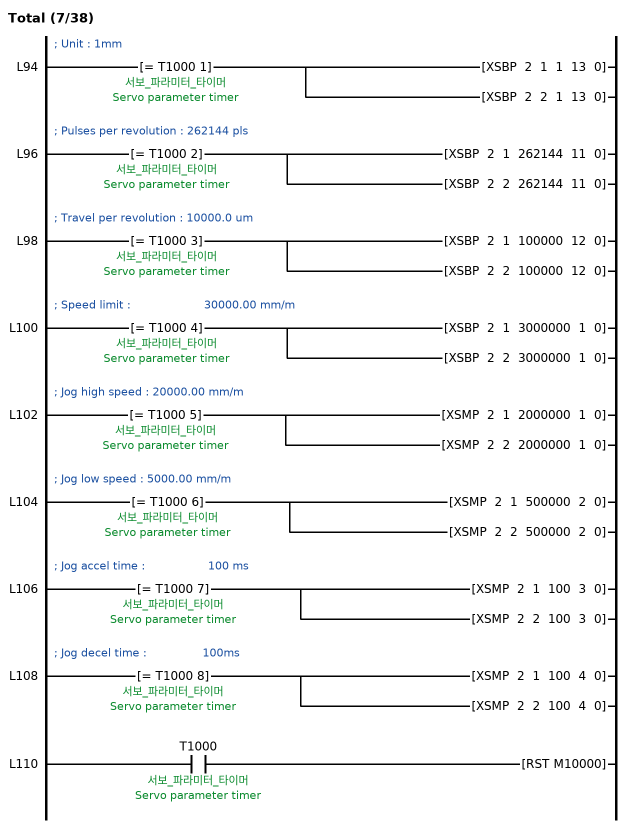
[picture p48: Total rungs L94-L110]
; L94
LOAD=     T1000 1	// 서보_파라미터_타이머 Servo parameter timer
XSBP      2 1 1 13 0
XSBP      2 2 1 13 0
// output comment: Unit : 1mm
; L96
LOAD=     T1000 2	// 서보_파라미터_타이머 Servo parameter timer
XSBP      2 1 262144 11 0
XSBP      2 2 262144 11 0
// output comment: Pulses per revolution : 262144 pls
; L98
LOAD=     T1000 3	// 서보_파라미터_타이머 Servo parameter timer
XSBP      2 1 100000 12 0
XSBP      2 2 100000 12 0
// output comment: Travel per revolution : 10000.0 um
; L100
LOAD=     T1000 4	// 서보_파라미터_타이머 Servo parameter timer
XSBP      2 1 3000000 1 0
XSBP      2 2 3000000 1 0
// output comment: Speed limit :                     30000.00 mm/m
; L102
LOAD=     T1000 5	// 서보_파라미터_타이머 Servo parameter timer
XSMP      2 1 2000000 1 0
XSMP      2 2 2000000 1 0
// output comment: Jog high speed : 20000.00 mm/m
; L104
LOAD=     T1000 6	// 서보_파라미터_타이머 Servo parameter timer
XSMP      2 1 500000 2 0
XSMP      2 2 500000 2 0
// output comment: Jog low speed : 5000.00 mm/m
; L106
LOAD=     T1000 7	// 서보_파라미터_타이머 Servo parameter timer
XSMP      2 1 100 3 0
XSMP      2 2 100 3 0
// output comment: Jog accel time :                  100 ms
; L108
LOAD=     T1000 8	// 서보_파라미터_타이머 Servo parameter timer
XSMP      2 1 100 4 0
XSMP      2 2 100 4 0
// output comment: Jog decel time :                100ms
; L110
LOAD      T1000	// 서보_파라미터_타이머 Servo parameter timer
RST       M10000

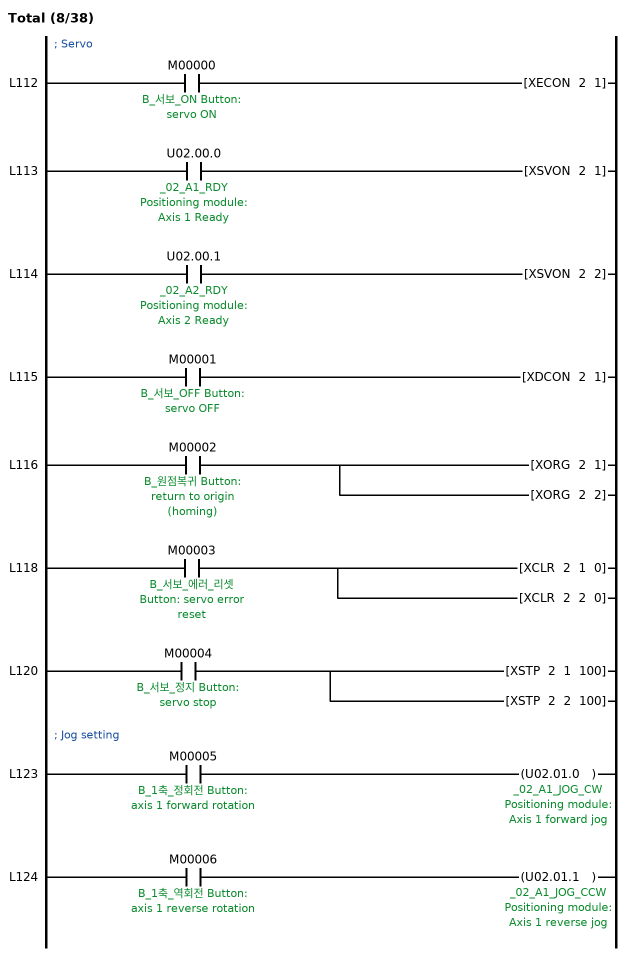
// Servo
; L112
LOAD      M00000	// B_서보_ON Button: servo ON
XECON     2 1
; L113
LOAD      U02.00.0	// _02_A1_RDY Positioning module: Axis 1 Ready
XSVON     2 1
; L114
LOAD      U02.00.1	// _02_A2_RDY Positioning module: Axis 2 Ready
XSVON     2 2
; L115
LOAD      M00001	// B_서보_OFF Button: servo OFF
XDCON     2 1
; L116
LOAD      M00002	// B_원점복귀 Button: return to origin (homing)
XORG      2 1
XORG      2 2
; L118
LOAD      M00003	// B_서보_에러_리셋 Button: servo error reset
XCLR      2 1 0
XCLR      2 2 0
; L120
LOAD      M00004	// B_서보_정지 Button: servo stop
XSTP      2 1 100
XSTP      2 2 100
// Jog setting
; L123
LOAD      M00005	// B_1축_정회전 Button: axis 1 forward rotation
OUT       U02.01.0	// _02_A1_JOG_CW Positioning module: Axis 1 forward jog
; L124
LOAD      M00006	// B_1축_역회전 Button: axis 1 reverse rotation
OUT       U02.01.1	// _02_A1_JOG_CCW Positioning module: Axis 1 reverse jog

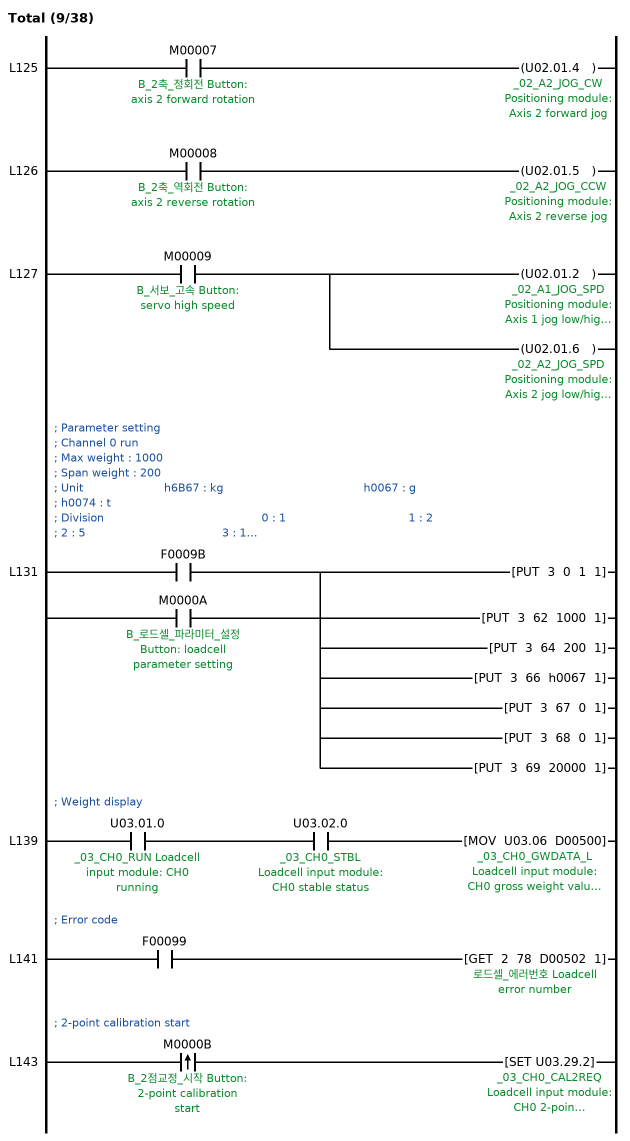
; L125
LOAD      M00007	// B_2축_정회전 Button: axis 2 forward rotation
OUT       U02.01.4	// _02_A2_JOG_CW Positioning module: Axis 2 forward jog
; L126
LOAD      M00008	// B_2축_역회전 Button: axis 2 reverse rotation
OUT       U02.01.5	// _02_A2_JOG_CCW Positioning module: Axis 2 reverse jog
; L127
LOAD      M00009	// B_서보_고속 Button: servo high speed
OUT       U02.01.2	// _02_A1_JOG_SPD Positioning module: Axis 1 jog low/high speed
OUT       U02.01.6	// _02_A2_JOG_SPD Positioning module: Axis 2 jog low/high speed
// Parameter setting
; L131
LOAD      F0009B
OR        M0000A	// B_로드셀_파라미터_설정 Button: loadcell parameter setting
PUT       3 0 1 1
PUT       3 62 1000 1
PUT       3 64 200 1
PUT       3 66 h0067 1
PUT       3 67 0 1
PUT       3 68 0 1
PUT       3 69 20000 1
// output comment: Channel 0 run
// output comment: Max weight : 1000
// output comment: Span weight : 200
// output comment: Unit                       h6B67 : kg                                        h0067 : g                                         h0074 : t
// output comment: Division                                             0 : 1                                   1 : 2                                             2 : 5                                       3 : 10
// output comment: Decimal                    0 : 1                    1: 0.1                         2 : 0.01                  3 : 0.001
// output comment: Loadcell sensitivity : 2mV/V
// Weight display
; L139
LOAD      U03.01.0	// _03_CH0_RUN Loadcell input module: CH0 running
AND       U03.02.0	// _03_CH0_STBL Loadcell input module: CH0 stable status
MOV       U03.06 D00500	// _03_CH0_GWDATA_L Loadcell input module: CH0 gross weight value (low) / Mass
// Error code
; L141
LOAD      F00099
GET       2 78 D00502 1	// 로드셀_에러번호 Loadcell error number
// 2-point calibration start
; L143
LOADP     M0000B	// B_2점교정_시작 Button: 2-point calibration start
SET       U03.29.2	// _03_CH0_CAL2REQ Loadcell input module: CH0 2-point calibration mode request

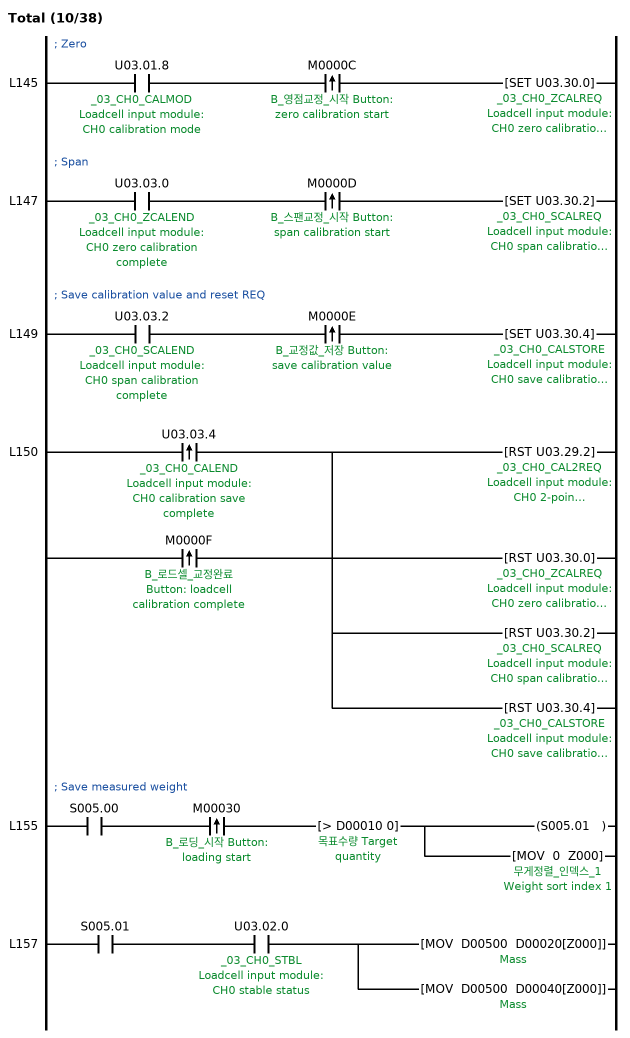
// Zero
; L145
LOAD      U03.01.8	// _03_CH0_CALMOD Loadcell input module: CH0 calibration mode
ANDP      M0000C	// B_영점교정_시작 Button: zero calibration start
SET       U03.30.0	// _03_CH0_ZCALREQ Loadcell input module: CH0 zero calibration command
// Span
; L147
LOAD      U03.03.0	// _03_CH0_ZCALEND Loadcell input module: CH0 zero calibration complete
ANDP      M0000D	// B_스팬교정_시작 Button: span calibration start
SET       U03.30.2	// _03_CH0_SCALREQ Loadcell input module: CH0 span calibration command
// Save calibration value and reset REQ
; L149
LOAD      U03.03.2	// _03_CH0_SCALEND Loadcell input module: CH0 span calibration complete
ANDP      M0000E	// B_교정값_저장 Button: save calibration value
SET       U03.30.4	// _03_CH0_CALSTORE Loadcell input module: CH0 save calibration value command
; L150
LOADP     U03.03.4	// _03_CH0_CALEND Loadcell input module: CH0 calibration save complete
ORP       M0000F	// B_로드셀_교정완료 Button: loadcell calibration complete
RST       U03.29.2	// _03_CH0_CAL2REQ Loadcell input module: CH0 2-point calibration mode request
RST       U03.30.0	// _03_CH0_ZCALREQ Loadcell input module: CH0 zero calibration command
RST       U03.30.2	// _03_CH0_SCALREQ Loadcell input module: CH0 span calibration command
RST       U03.30.4	// _03_CH0_CALSTORE Loadcell input module: CH0 save calibration value command
// Save measured weight
; L155
LOAD      S005.00
ANDP      M00030	// B_로딩_시작 Button: loading start
AND>      D00010 0	// 목표수량 Target quantity
OUT       S005.01
MOV       0 Z000	// 무게정렬_인덱스_1 Weight sort index 1
; L157
LOAD      S005.01
AND       U03.02.0	// _03_CH0_STBL Loadcell input module: CH0 stable status
MOV       D00500 D00020[Z000]	// Mass
MOV       D00500 D00040[Z000]	// Mass

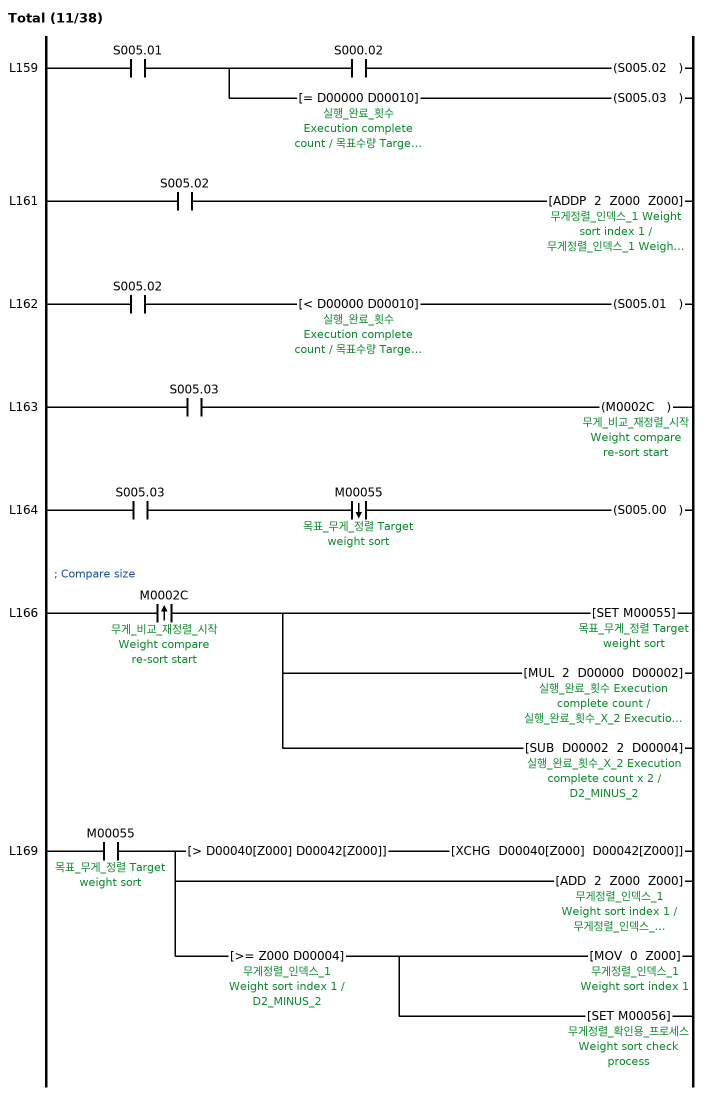
; L159
LOAD      S005.01
MPUSH
AND       S000.02
OUT       S005.02
MPOP
AND=      D00000 D00010	// 실행_완료_횟수 Execution complete count / 목표수량 Target quantity
OUT       S005.03
; L161
LOAD      S005.02
ADDP      2 Z000 Z000	// 무게정렬_인덱스_1 Weight sort index 1 / 무게정렬_인덱스_1 Weight sort index 1
; L162
LOAD      S005.02
AND<      D00000 D00010	// 실행_완료_횟수 Execution complete count / 목표수량 Target quantity
OUT       S005.01
; L163
LOAD      S005.03
OUT       M0002C	// 무게_비교_재정렬_시작 Weight compare re-sort start
; L164
LOAD      S005.03
ANDN      M00055	// 목표_무게_정렬 Target weight sort
OUT       S005.00
// Compare size
; L166
LOADP     M0002C	// 무게_비교_재정렬_시작 Weight compare re-sort start
SET       M00055	// 목표_무게_정렬 Target weight sort
MUL       2 D00000 D00002	// 실행_완료_횟수 Execution complete count / 실행_완료_횟수_X_2 Execution complete count x 2
SUB       D00002 2 D00004	// 실행_완료_횟수_X_2 Execution complete count x 2 / D2_MINUS_2
; L169
LOAD      M00055	// 목표_무게_정렬 Target weight sort
MPUSH
AND>      D00040[Z000] D00042[Z000]
XCHG      D00040[Z000] D00042[Z000]
MPOP
ADD       2 Z000 Z000	// 무게정렬_인덱스_1 Weight sort index 1 / 무게정렬_인덱스_1 Weight sort index 1
AND>=     Z000 D00004	// 무게정렬_인덱스_1 Weight sort index 1 / D2_MINUS_2
MOV       0 Z000	// 무게정렬_인덱스_1 Weight sort index 1
SET       M00056	// 무게정렬_확인용_프로세스 Weight sort check process

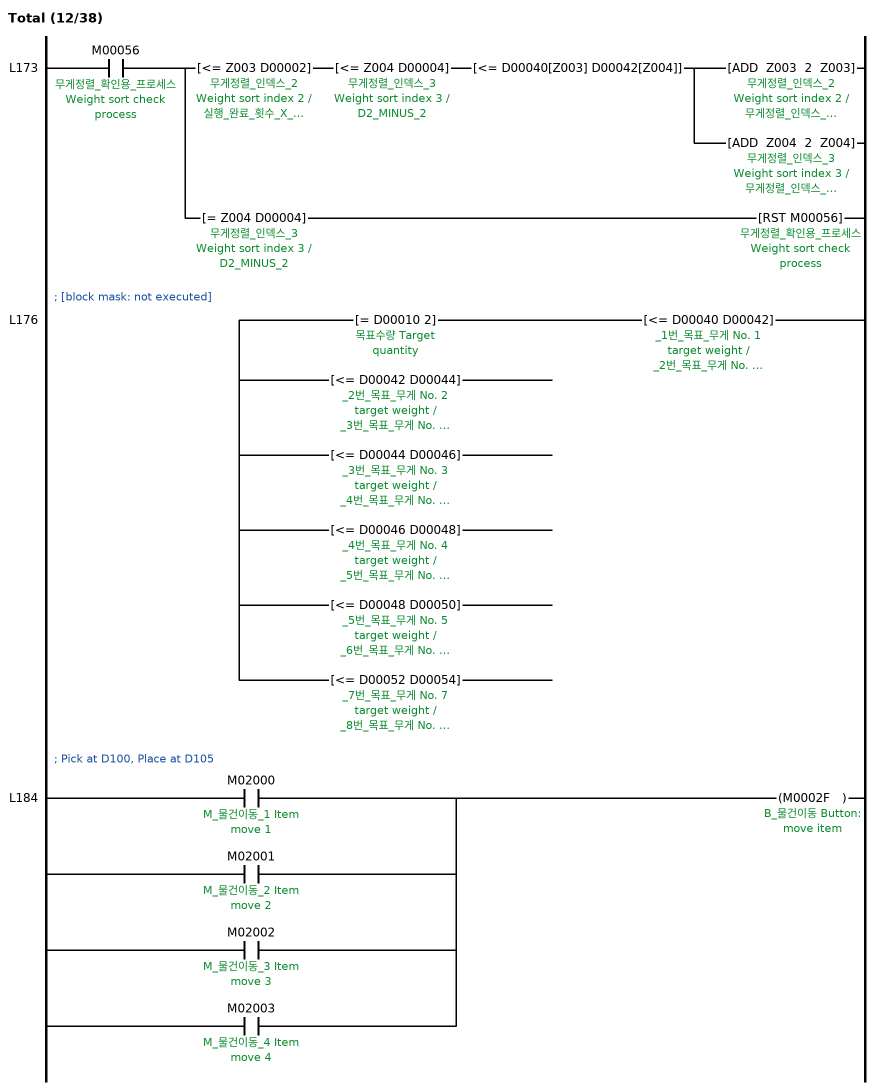
; L173
LOAD      M00056	// 무게정렬_확인용_프로세스 Weight sort check process
MPUSH
AND<=     Z003 D00002	// 무게정렬_인덱스_2 Weight sort index 2 / 실행_완료_횟수_X_2 Execution complete count x 2
AND<=     Z004 D00004	// 무게정렬_인덱스_3 Weight sort index 3 / D2_MINUS_2
AND<=     D00040[Z003] D00042[Z004]
ADD       Z003 2 Z003	// 무게정렬_인덱스_2 Weight sort index 2 / 무게정렬_인덱스_2 Weight sort index 2
ADD       Z004 2 Z004	// 무게정렬_인덱스_3 Weight sort index 3 / 무게정렬_인덱스_3 Weight sort index 3
MPOP
AND=      Z004 D00004	// 무게정렬_인덱스_3 Weight sort index 3 / D2_MINUS_2
RST       M00056	// 무게정렬_확인용_프로세스 Weight sort check process
; L176 (block mask: not executed)
// network not rendered as a mnemonic list; see the picture
// Pick at D100, Place at D105
; L184
LOAD      M02000	// M_물건이동_1 Item move 1
OR        M02001	// M_물건이동_2 Item move 2
OR        M02002	// M_물건이동_3 Item move 3
OR        M02003	// M_물건이동_4 Item move 4
OUT       M0002F	// B_물건이동 Button: move item

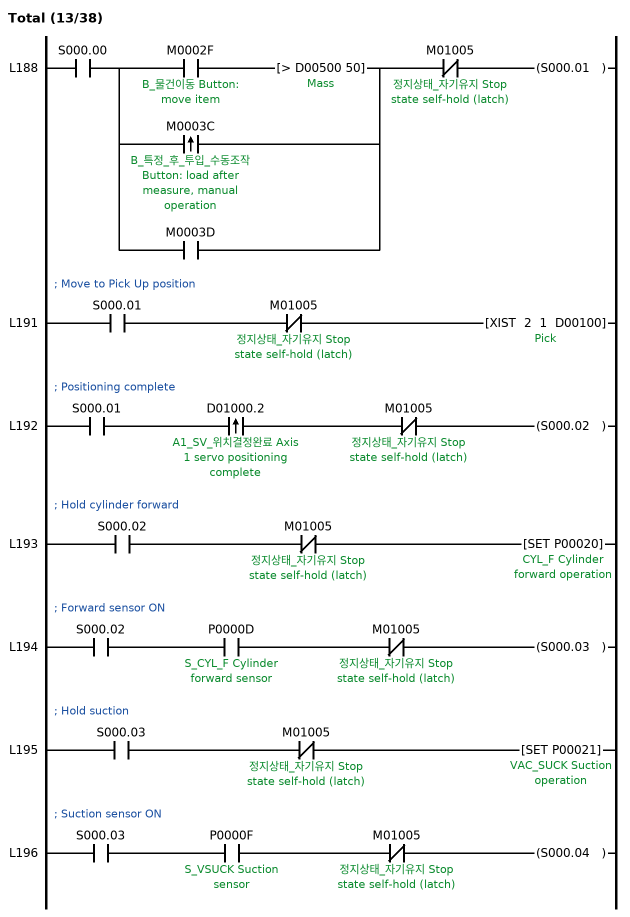
; L188
LOAD      S000.00
LOAD      M0002F	// B_물건이동 Button: move item
AND>      D00500 50	// Mass
ORP       M0003C	// B_특정_후_투입_수동조작 Button: load after measure, manual operation
OR        M0003D
AND LOAD
AND NOT   M01005	// 정지상태_자기유지 Stop state self-hold (latch)
OUT       S000.01
; L191
LOAD      S000.01
AND NOT   M01005	// 정지상태_자기유지 Stop state self-hold (latch)
XIST      2 1 D00100	// Pick
// output comment: Move to Pick Up position
; L192
LOAD      S000.01
ANDP      D01000.2	// A1_SV_위치결정완료 Axis 1 servo positioning complete
AND NOT   M01005	// 정지상태_자기유지 Stop state self-hold (latch)
OUT       S000.02
// output comment: Positioning complete
; L193
LOAD      S000.02
AND NOT   M01005	// 정지상태_자기유지 Stop state self-hold (latch)
SET       P00020	// CYL_F Cylinder forward operation
// output comment: Hold cylinder forward
; L194
LOAD      S000.02
AND       P0000D	// S_CYL_F Cylinder forward sensor
AND NOT   M01005	// 정지상태_자기유지 Stop state self-hold (latch)
OUT       S000.03
// output comment: Forward sensor ON
; L195
LOAD      S000.03
AND NOT   M01005	// 정지상태_자기유지 Stop state self-hold (latch)
SET       P00021	// VAC_SUCK Suction operation
// output comment: Hold suction
; L196
LOAD      S000.03
AND       P0000F	// S_VSUCK Suction sensor
AND NOT   M01005	// 정지상태_자기유지 Stop state self-hold (latch)
OUT       S000.04
// output comment: Suction sensor ON

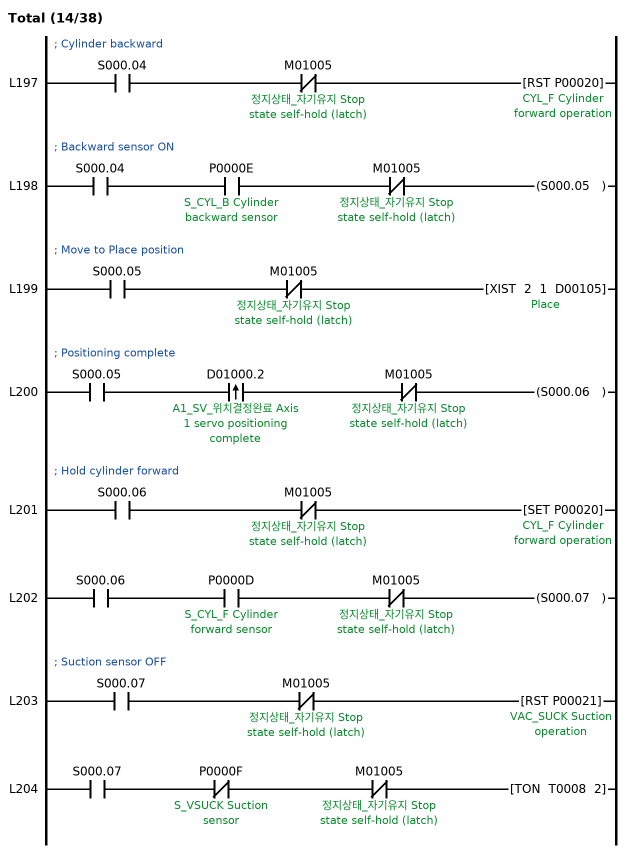
; L197
LOAD      S000.04
AND NOT   M01005	// 정지상태_자기유지 Stop state self-hold (latch)
RST       P00020	// CYL_F Cylinder forward operation
// output comment: Cylinder backward
; L198
LOAD      S000.04
AND       P0000E	// S_CYL_B Cylinder backward sensor
AND NOT   M01005	// 정지상태_자기유지 Stop state self-hold (latch)
OUT       S000.05
// output comment: Backward sensor ON
; L199
LOAD      S000.05
AND NOT   M01005	// 정지상태_자기유지 Stop state self-hold (latch)
XIST      2 1 D00105	// Place
// output comment: Move to Place position
; L200
LOAD      S000.05
ANDP      D01000.2	// A1_SV_위치결정완료 Axis 1 servo positioning complete
AND NOT   M01005	// 정지상태_자기유지 Stop state self-hold (latch)
OUT       S000.06
// output comment: Positioning complete
; L201
LOAD      S000.06
AND NOT   M01005	// 정지상태_자기유지 Stop state self-hold (latch)
SET       P00020	// CYL_F Cylinder forward operation
// output comment: Hold cylinder forward
; L202
LOAD      S000.06
AND       P0000D	// S_CYL_F Cylinder forward sensor
AND NOT   M01005	// 정지상태_자기유지 Stop state self-hold (latch)
OUT       S000.07
; L203
LOAD      S000.07
AND NOT   M01005	// 정지상태_자기유지 Stop state self-hold (latch)
RST       P00021	// VAC_SUCK Suction operation
// output comment: Suction sensor OFF
; L204
LOAD      S000.07
AND NOT   P0000F	// S_VSUCK Suction sensor
AND NOT   M01005	// 정지상태_자기유지 Stop state self-hold (latch)
TON       T0008 2

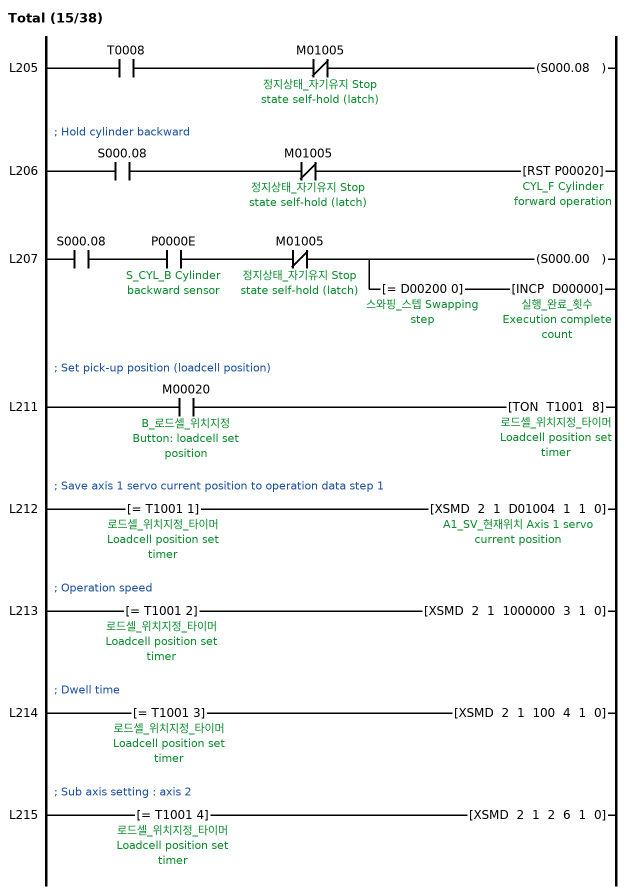
; L205
LOAD      T0008
AND NOT   M01005	// 정지상태_자기유지 Stop state self-hold (latch)
OUT       S000.08
; L206
LOAD      S000.08
AND NOT   M01005	// 정지상태_자기유지 Stop state self-hold (latch)
RST       P00020	// CYL_F Cylinder forward operation
// output comment: Hold cylinder backward
; L207
LOAD      S000.08
AND       P0000E	// S_CYL_B Cylinder backward sensor
AND NOT   M01005	// 정지상태_자기유지 Stop state self-hold (latch)
OUT       S000.00
AND=      D00200 0	// 스와핑_스텝 Swapping step
INCP      D00000	// 실행_완료_횟수 Execution complete count
// Set pick-up position (loadcell position)
; L211
LOAD      M00020	// B_로드셀_위치지정 Button: loadcell set position
TON       T1001 8	// 로드셀_위치지정_타이머 Loadcell position set timer
; L212
LOAD=     T1001 1	// 로드셀_위치지정_타이머 Loadcell position set timer
XSMD      2 1 D01004 1 1 0	// A1_SV_현재위치 Axis 1 servo current position
// output comment: Save axis 1 servo current position to operation data step 1
; L213
LOAD=     T1001 2	// 로드셀_위치지정_타이머 Loadcell position set timer
XSMD      2 1 1000000 3 1 0
// output comment: Operation speed
; L214
LOAD=     T1001 3	// 로드셀_위치지정_타이머 Loadcell position set timer
XSMD      2 1 100 4 1 0
// output comment: Dwell time
; L215
LOAD=     T1001 4	// 로드셀_위치지정_타이머 Loadcell position set timer
XSMD      2 1 2 6 1 0
// output comment: Sub axis setting : axis 2

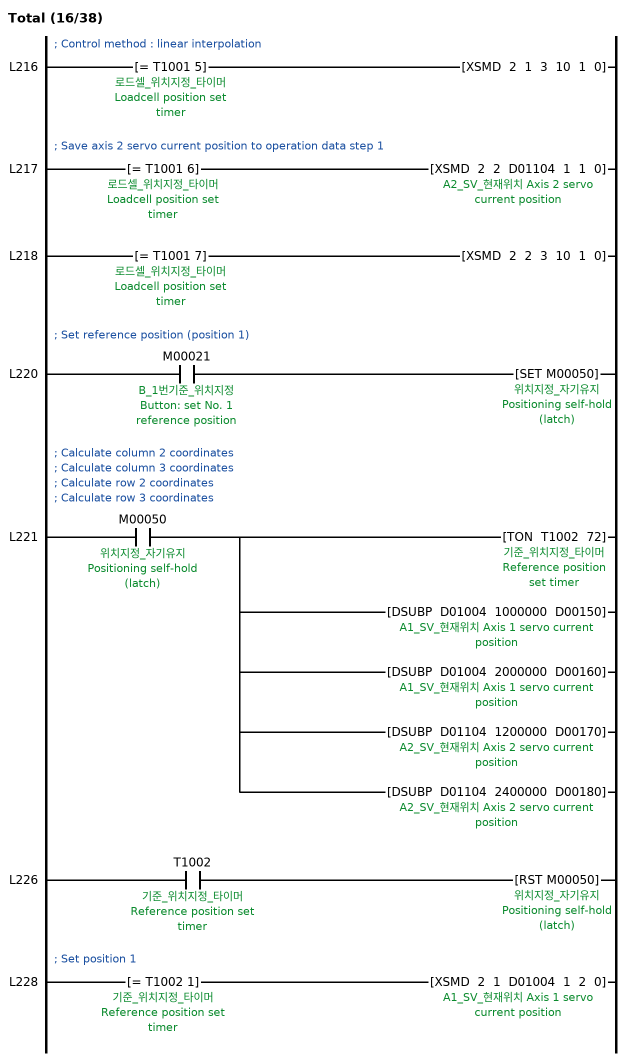
; L216
LOAD=     T1001 5	// 로드셀_위치지정_타이머 Loadcell position set timer
XSMD      2 1 3 10 1 0
// output comment: Control method : linear interpolation
; L217
LOAD=     T1001 6	// 로드셀_위치지정_타이머 Loadcell position set timer
XSMD      2 2 D01104 1 1 0	// A2_SV_현재위치 Axis 2 servo current position
// output comment: Save axis 2 servo current position to operation data step 1
; L218
LOAD=     T1001 7	// 로드셀_위치지정_타이머 Loadcell position set timer
XSMD      2 2 3 10 1 0
// output comment: 
// Set reference position (position 1)
; L220
LOAD      M00021	// B_1번기준_위치지정 Button: set No. 1 reference position
SET       M00050	// 위치지정_자기유지 Positioning self-hold (latch)
; L221
LOAD      M00050	// 위치지정_자기유지 Positioning self-hold (latch)
TON       T1002 72	// 기준_위치지정_타이머 Reference position set timer
DSUBP     D01004 1000000 D00150	// A1_SV_현재위치 Axis 1 servo current position
DSUBP     D01004 2000000 D00160	// A1_SV_현재위치 Axis 1 servo current position
DSUBP     D01104 1200000 D00170	// A2_SV_현재위치 Axis 2 servo current position
DSUBP     D01104 2400000 D00180	// A2_SV_현재위치 Axis 2 servo current position
// output comment: Calculate column 2 coordinates
// output comment: Calculate column 3 coordinates
// output comment: Calculate row 2 coordinates
// output comment: Calculate row 3 coordinates
; L226
LOAD      T1002	// 기준_위치지정_타이머 Reference position set timer
RST       M00050	// 위치지정_자기유지 Positioning self-hold (latch)
// Set position 1
; L228
LOAD=     T1002 1	// 기준_위치지정_타이머 Reference position set timer
XSMD      2 1 D01004 1 2 0	// A1_SV_현재위치 Axis 1 servo current position

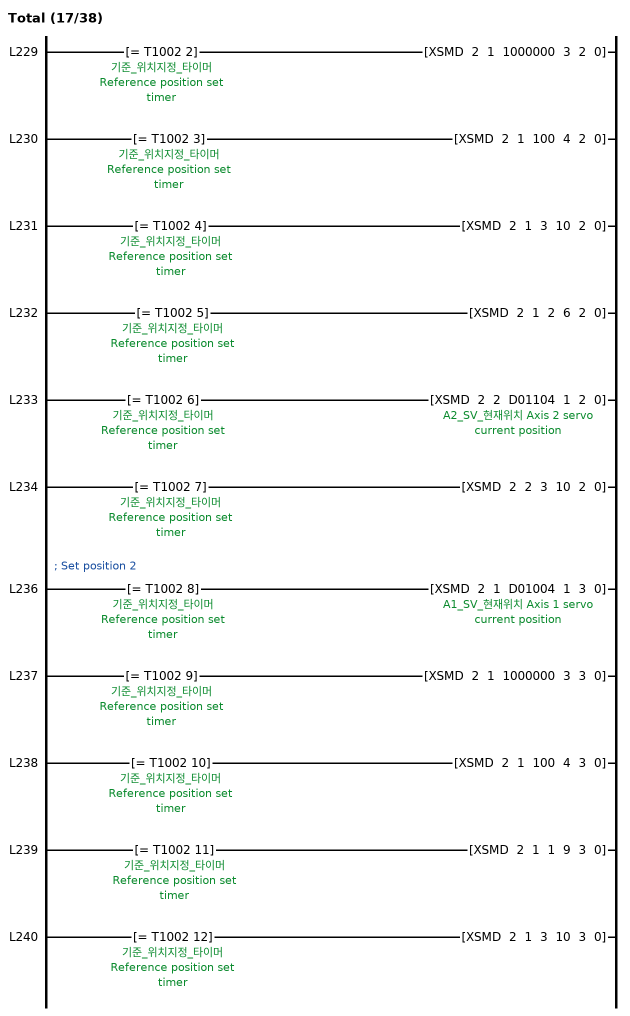
; L229
LOAD=     T1002 2	// 기준_위치지정_타이머 Reference position set timer
XSMD      2 1 1000000 3 2 0
; L230
LOAD=     T1002 3	// 기준_위치지정_타이머 Reference position set timer
XSMD      2 1 100 4 2 0
; L231
LOAD=     T1002 4	// 기준_위치지정_타이머 Reference position set timer
XSMD      2 1 3 10 2 0
; L232
LOAD=     T1002 5	// 기준_위치지정_타이머 Reference position set timer
XSMD      2 1 2 6 2 0
; L233
LOAD=     T1002 6	// 기준_위치지정_타이머 Reference position set timer
XSMD      2 2 D01104 1 2 0	// A2_SV_현재위치 Axis 2 servo current position
; L234
LOAD=     T1002 7	// 기준_위치지정_타이머 Reference position set timer
XSMD      2 2 3 10 2 0
// Set position 2
; L236
LOAD=     T1002 8	// 기준_위치지정_타이머 Reference position set timer
XSMD      2 1 D01004 1 3 0	// A1_SV_현재위치 Axis 1 servo current position
; L237
LOAD=     T1002 9	// 기준_위치지정_타이머 Reference position set timer
XSMD      2 1 1000000 3 3 0
; L238
LOAD=     T1002 10	// 기준_위치지정_타이머 Reference position set timer
XSMD      2 1 100 4 3 0
; L239
LOAD=     T1002 11	// 기준_위치지정_타이머 Reference position set timer
XSMD      2 1 1 9 3 0
; L240
LOAD=     T1002 12	// 기준_위치지정_타이머 Reference position set timer
XSMD      2 1 3 10 3 0

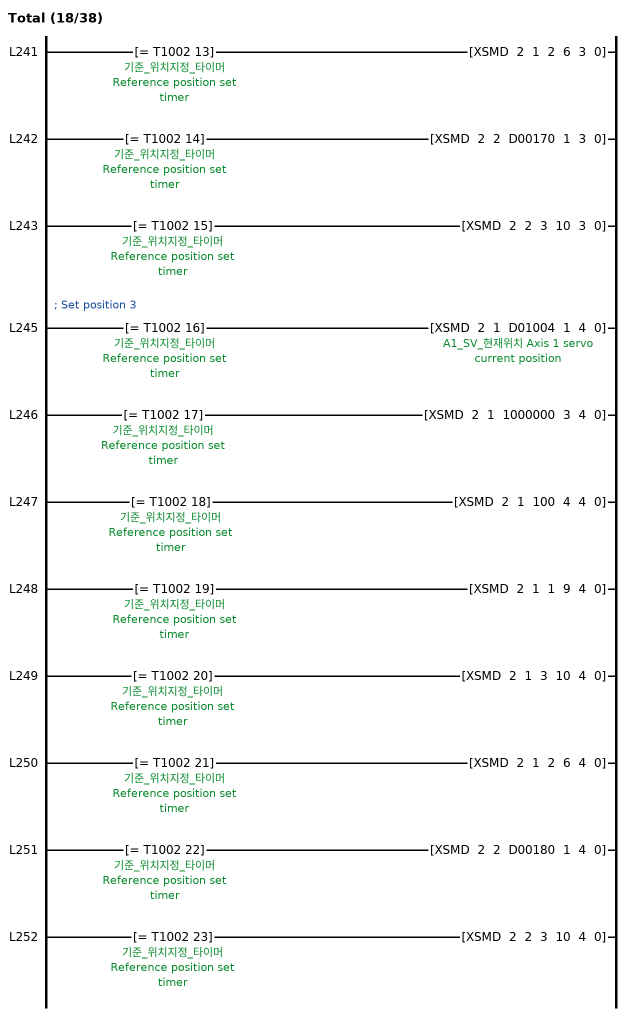
; L241
LOAD=     T1002 13	// 기준_위치지정_타이머 Reference position set timer
XSMD      2 1 2 6 3 0
; L242
LOAD=     T1002 14	// 기준_위치지정_타이머 Reference position set timer
XSMD      2 2 D00170 1 3 0
; L243
LOAD=     T1002 15	// 기준_위치지정_타이머 Reference position set timer
XSMD      2 2 3 10 3 0
// Set position 3
; L245
LOAD=     T1002 16	// 기준_위치지정_타이머 Reference position set timer
XSMD      2 1 D01004 1 4 0	// A1_SV_현재위치 Axis 1 servo current position
; L246
LOAD=     T1002 17	// 기준_위치지정_타이머 Reference position set timer
XSMD      2 1 1000000 3 4 0
; L247
LOAD=     T1002 18	// 기준_위치지정_타이머 Reference position set timer
XSMD      2 1 100 4 4 0
; L248
LOAD=     T1002 19	// 기준_위치지정_타이머 Reference position set timer
XSMD      2 1 1 9 4 0
; L249
LOAD=     T1002 20	// 기준_위치지정_타이머 Reference position set timer
XSMD      2 1 3 10 4 0
; L250
LOAD=     T1002 21	// 기준_위치지정_타이머 Reference position set timer
XSMD      2 1 2 6 4 0
; L251
LOAD=     T1002 22	// 기준_위치지정_타이머 Reference position set timer
XSMD      2 2 D00180 1 4 0
; L252
LOAD=     T1002 23	// 기준_위치지정_타이머 Reference position set timer
XSMD      2 2 3 10 4 0

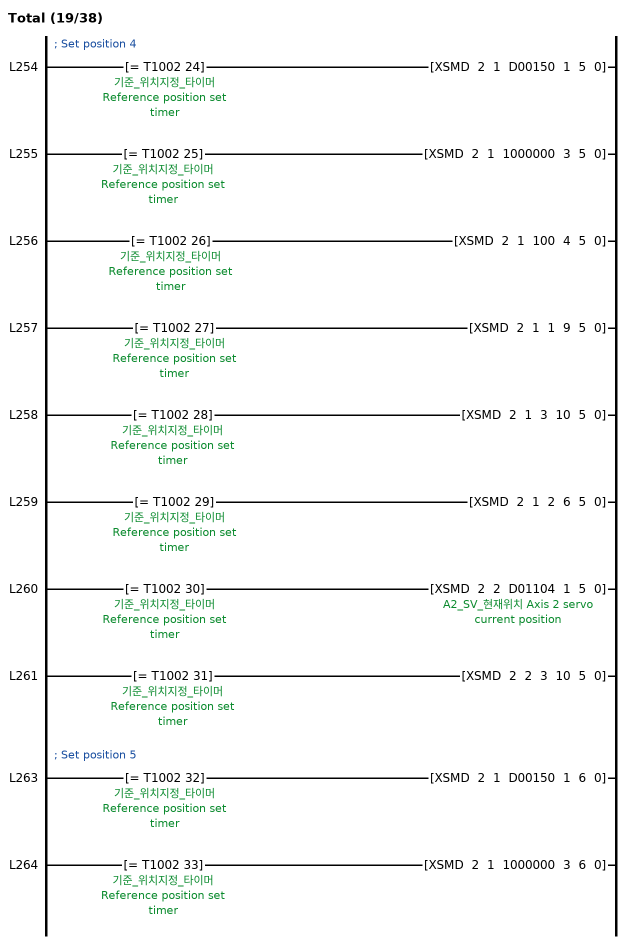
// Set position 4
; L254
LOAD=     T1002 24	// 기준_위치지정_타이머 Reference position set timer
XSMD      2 1 D00150 1 5 0
; L255
LOAD=     T1002 25	// 기준_위치지정_타이머 Reference position set timer
XSMD      2 1 1000000 3 5 0
; L256
LOAD=     T1002 26	// 기준_위치지정_타이머 Reference position set timer
XSMD      2 1 100 4 5 0
; L257
LOAD=     T1002 27	// 기준_위치지정_타이머 Reference position set timer
XSMD      2 1 1 9 5 0
; L258
LOAD=     T1002 28	// 기준_위치지정_타이머 Reference position set timer
XSMD      2 1 3 10 5 0
; L259
LOAD=     T1002 29	// 기준_위치지정_타이머 Reference position set timer
XSMD      2 1 2 6 5 0
; L260
LOAD=     T1002 30	// 기준_위치지정_타이머 Reference position set timer
XSMD      2 2 D01104 1 5 0	// A2_SV_현재위치 Axis 2 servo current position
; L261
LOAD=     T1002 31	// 기준_위치지정_타이머 Reference position set timer
XSMD      2 2 3 10 5 0
// Set position 5
; L263
LOAD=     T1002 32	// 기준_위치지정_타이머 Reference position set timer
XSMD      2 1 D00150 1 6 0
; L264
LOAD=     T1002 33	// 기준_위치지정_타이머 Reference position set timer
XSMD      2 1 1000000 3 6 0

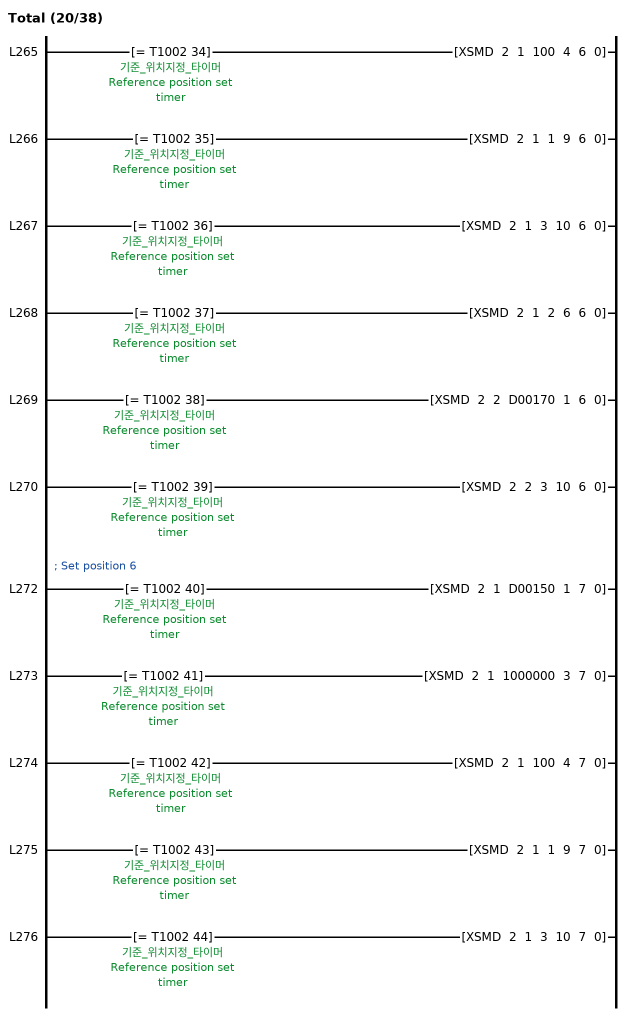
; L265
LOAD=     T1002 34	// 기준_위치지정_타이머 Reference position set timer
XSMD      2 1 100 4 6 0
; L266
LOAD=     T1002 35	// 기준_위치지정_타이머 Reference position set timer
XSMD      2 1 1 9 6 0
; L267
LOAD=     T1002 36	// 기준_위치지정_타이머 Reference position set timer
XSMD      2 1 3 10 6 0
; L268
LOAD=     T1002 37	// 기준_위치지정_타이머 Reference position set timer
XSMD      2 1 2 6 6 0
; L269
LOAD=     T1002 38	// 기준_위치지정_타이머 Reference position set timer
XSMD      2 2 D00170 1 6 0
; L270
LOAD=     T1002 39	// 기준_위치지정_타이머 Reference position set timer
XSMD      2 2 3 10 6 0
// Set position 6
; L272
LOAD=     T1002 40	// 기준_위치지정_타이머 Reference position set timer
XSMD      2 1 D00150 1 7 0
; L273
LOAD=     T1002 41	// 기준_위치지정_타이머 Reference position set timer
XSMD      2 1 1000000 3 7 0
; L274
LOAD=     T1002 42	// 기준_위치지정_타이머 Reference position set timer
XSMD      2 1 100 4 7 0
; L275
LOAD=     T1002 43	// 기준_위치지정_타이머 Reference position set timer
XSMD      2 1 1 9 7 0
; L276
LOAD=     T1002 44	// 기준_위치지정_타이머 Reference position set timer
XSMD      2 1 3 10 7 0

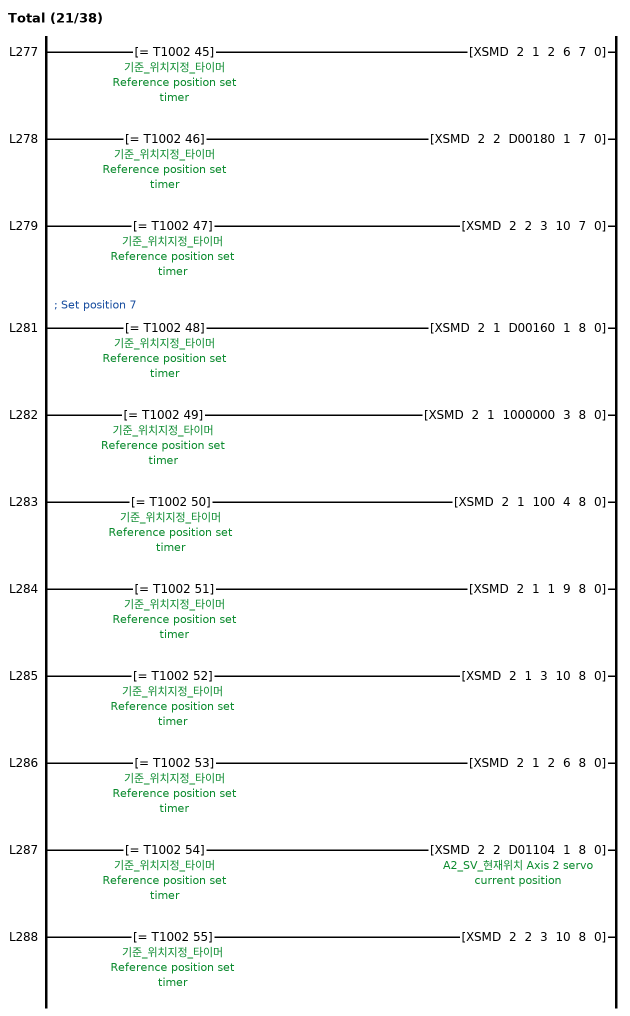
; L277
LOAD=     T1002 45	// 기준_위치지정_타이머 Reference position set timer
XSMD      2 1 2 6 7 0
; L278
LOAD=     T1002 46	// 기준_위치지정_타이머 Reference position set timer
XSMD      2 2 D00180 1 7 0
; L279
LOAD=     T1002 47	// 기준_위치지정_타이머 Reference position set timer
XSMD      2 2 3 10 7 0
// Set position 7
; L281
LOAD=     T1002 48	// 기준_위치지정_타이머 Reference position set timer
XSMD      2 1 D00160 1 8 0
; L282
LOAD=     T1002 49	// 기준_위치지정_타이머 Reference position set timer
XSMD      2 1 1000000 3 8 0
; L283
LOAD=     T1002 50	// 기준_위치지정_타이머 Reference position set timer
XSMD      2 1 100 4 8 0
; L284
LOAD=     T1002 51	// 기준_위치지정_타이머 Reference position set timer
XSMD      2 1 1 9 8 0
; L285
LOAD=     T1002 52	// 기준_위치지정_타이머 Reference position set timer
XSMD      2 1 3 10 8 0
; L286
LOAD=     T1002 53	// 기준_위치지정_타이머 Reference position set timer
XSMD      2 1 2 6 8 0
; L287
LOAD=     T1002 54	// 기준_위치지정_타이머 Reference position set timer
XSMD      2 2 D01104 1 8 0	// A2_SV_현재위치 Axis 2 servo current position
; L288
LOAD=     T1002 55	// 기준_위치지정_타이머 Reference position set timer
XSMD      2 2 3 10 8 0

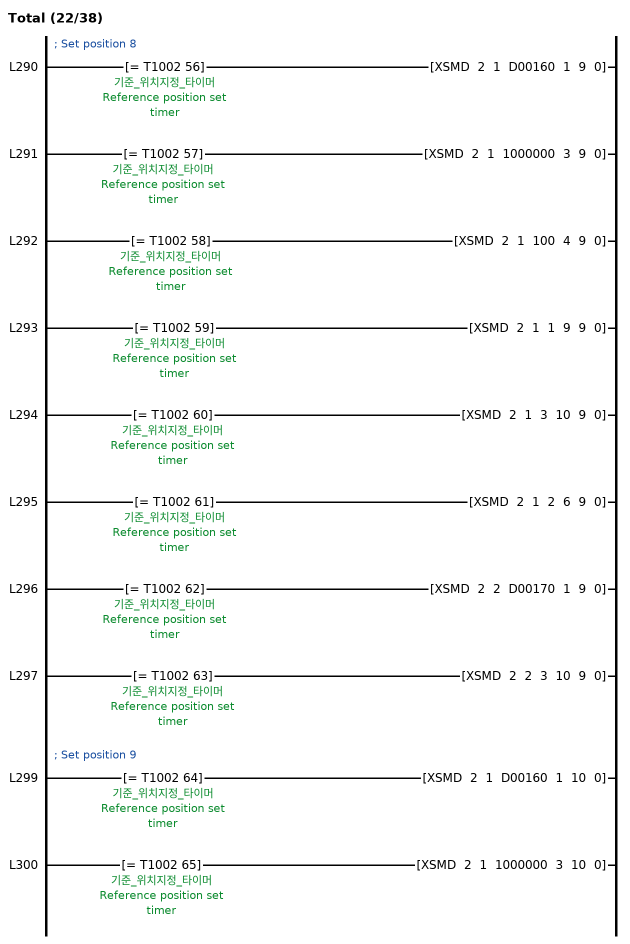
// Set position 8
; L290
LOAD=     T1002 56	// 기준_위치지정_타이머 Reference position set timer
XSMD      2 1 D00160 1 9 0
; L291
LOAD=     T1002 57	// 기준_위치지정_타이머 Reference position set timer
XSMD      2 1 1000000 3 9 0
; L292
LOAD=     T1002 58	// 기준_위치지정_타이머 Reference position set timer
XSMD      2 1 100 4 9 0
; L293
LOAD=     T1002 59	// 기준_위치지정_타이머 Reference position set timer
XSMD      2 1 1 9 9 0
; L294
LOAD=     T1002 60	// 기준_위치지정_타이머 Reference position set timer
XSMD      2 1 3 10 9 0
; L295
LOAD=     T1002 61	// 기준_위치지정_타이머 Reference position set timer
XSMD      2 1 2 6 9 0
; L296
LOAD=     T1002 62	// 기준_위치지정_타이머 Reference position set timer
XSMD      2 2 D00170 1 9 0
; L297
LOAD=     T1002 63	// 기준_위치지정_타이머 Reference position set timer
XSMD      2 2 3 10 9 0
// Set position 9
; L299
LOAD=     T1002 64	// 기준_위치지정_타이머 Reference position set timer
XSMD      2 1 D00160 1 10 0
; L300
LOAD=     T1002 65	// 기준_위치지정_타이머 Reference position set timer
XSMD      2 1 1000000 3 10 0

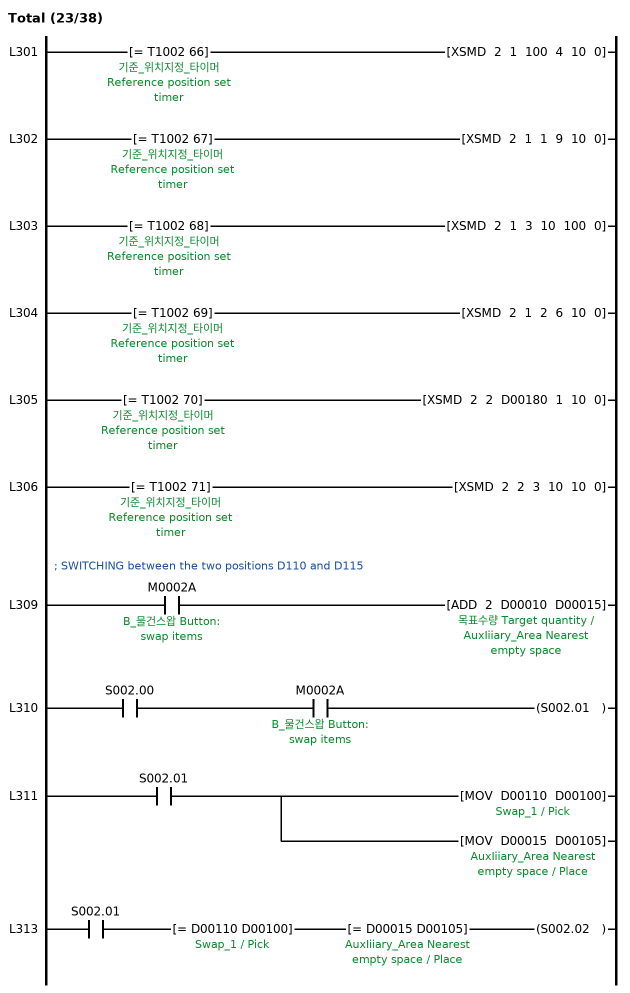
; L301
LOAD=     T1002 66	// 기준_위치지정_타이머 Reference position set timer
XSMD      2 1 100 4 10 0
; L302
LOAD=     T1002 67	// 기준_위치지정_타이머 Reference position set timer
XSMD      2 1 1 9 10 0
; L303
LOAD=     T1002 68	// 기준_위치지정_타이머 Reference position set timer
XSMD      2 1 3 10 100 0
; L304
LOAD=     T1002 69	// 기준_위치지정_타이머 Reference position set timer
XSMD      2 1 2 6 10 0
; L305
LOAD=     T1002 70	// 기준_위치지정_타이머 Reference position set timer
XSMD      2 2 D00180 1 10 0
; L306
LOAD=     T1002 71	// 기준_위치지정_타이머 Reference position set timer
XSMD      2 2 3 10 10 0
// SWITCHING between the two positions D110 and D115
; L309
LOAD      M0002A	// B_물건스왑 Button: swap items
ADD       2 D00010 D00015	// 목표수량 Target quantity / AuxIiiary_Area Nearest empty space
; L310
LOAD      S002.00
AND       M0002A	// B_물건스왑 Button: swap items
OUT       S002.01
; L311
LOAD      S002.01
MOV       D00110 D00100	// Swap_1 / Pick
MOV       D00015 D00105	// AuxIiiary_Area Nearest empty space / Place
; L313
LOAD      S002.01
AND=      D00110 D00100	// Swap_1 / Pick
AND=      D00015 D00105	// AuxIiiary_Area Nearest empty space / Place
OUT       S002.02

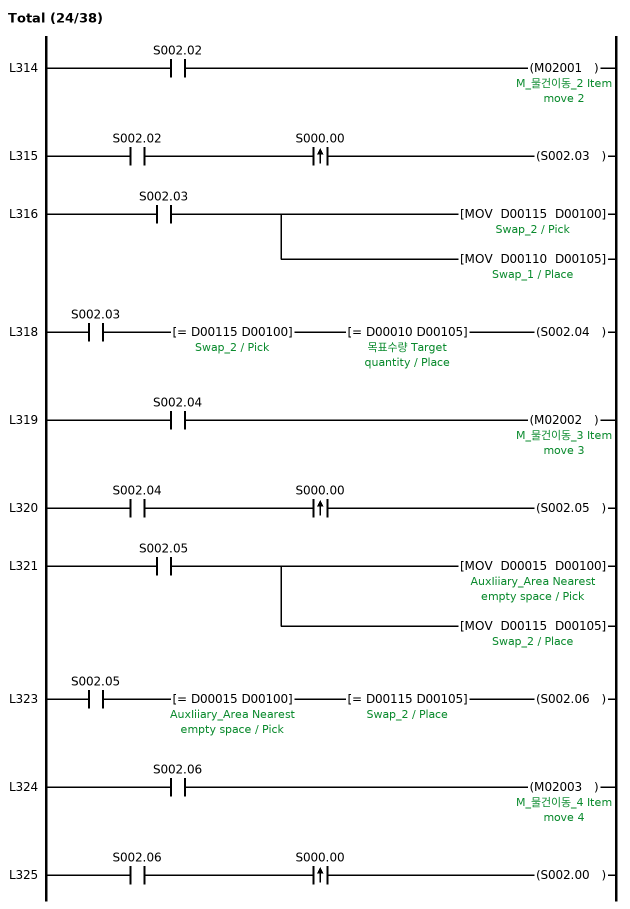
; L314
LOAD      S002.02
OUT       M02001	// M_물건이동_2 Item move 2
; L315
LOAD      S002.02
ANDP      S000.00
OUT       S002.03
; L316
LOAD      S002.03
MOV       D00115 D00100	// Swap_2 / Pick
MOV       D00110 D00105	// Swap_1 / Place
; L318
LOAD      S002.03
AND=      D00115 D00100	// Swap_2 / Pick
AND=      D00010 D00105	// 목표수량 Target quantity / Place
OUT       S002.04
; L319
LOAD      S002.04
OUT       M02002	// M_물건이동_3 Item move 3
; L320
LOAD      S002.04
ANDP      S000.00
OUT       S002.05
; L321
LOAD      S002.05
MOV       D00015 D00100	// AuxIiiary_Area Nearest empty space / Pick
MOV       D00115 D00105	// Swap_2 / Place
; L323
LOAD      S002.05
AND=      D00015 D00100	// AuxIiiary_Area Nearest empty space / Pick
AND=      D00115 D00105	// Swap_2 / Place
OUT       S002.06
; L324
LOAD      S002.06
OUT       M02003	// M_물건이동_4 Item move 4
; L325
LOAD      S002.06
ANDP      S000.00
OUT       S002.00

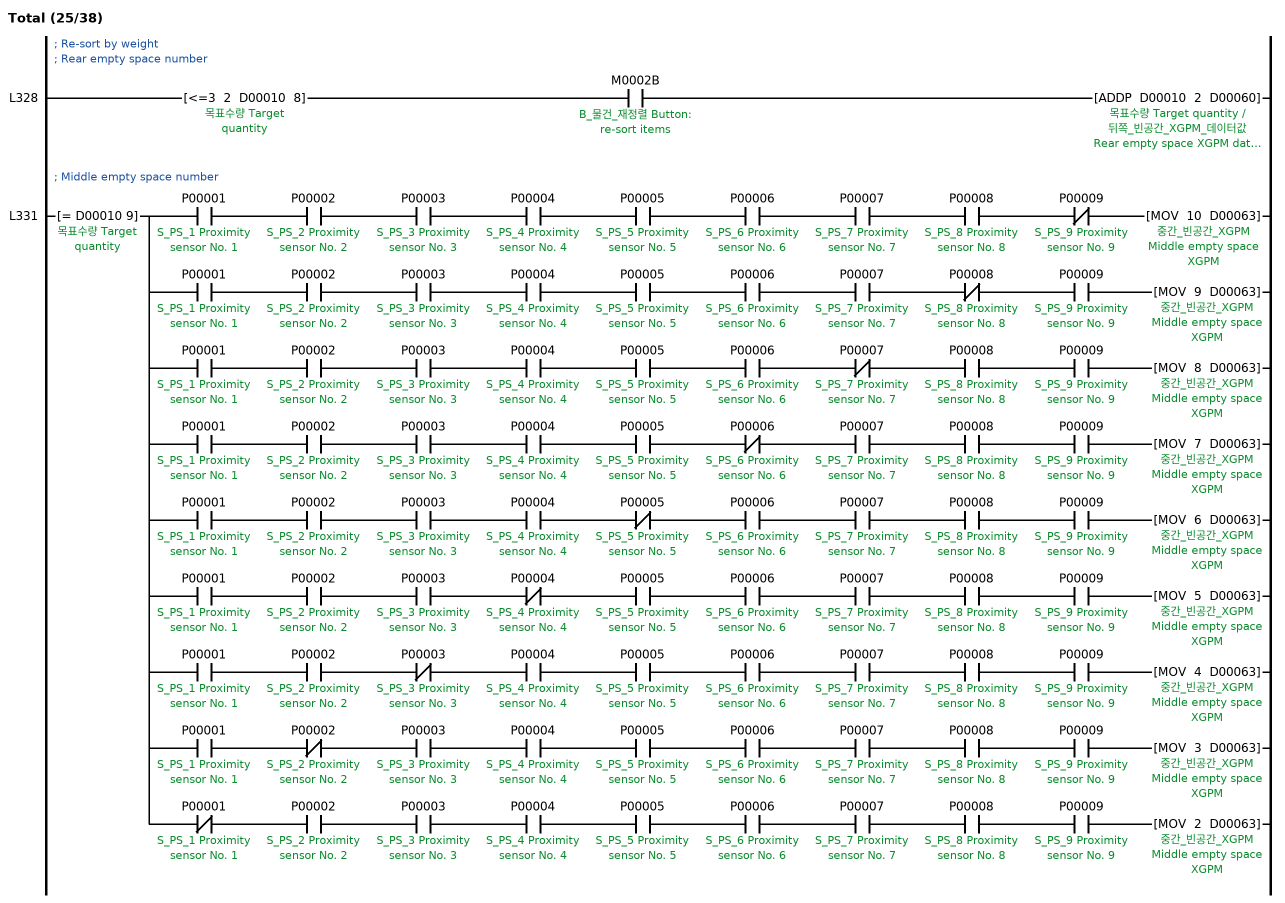
// Re-sort by weight
// Rear empty space number
; L328
LOAD<=3   2 D00010 8	// 목표수량 Target quantity
AND       M0002B	// B_물건_재정렬 Button: re-sort items
ADDP      D00010 2 D00060	// 목표수량 Target quantity / 뒤쪽_빈공간_XGPM_데이터값 Rear empty space XGPM data value
// Middle empty space number
; L331
LOAD=     D00010 9	// 목표수량 Target quantity
MPUSH
AND       P00001	// S_PS_1 Proximity sensor No. 1
AND       P00002	// S_PS_2 Proximity sensor No. 2
AND       P00003	// S_PS_3 Proximity sensor No. 3
AND       P00004	// S_PS_4 Proximity sensor No. 4
AND       P00005	// S_PS_5 Proximity sensor No. 5
AND       P00006	// S_PS_6 Proximity sensor No. 6
AND       P00007	// S_PS_7 Proximity sensor No. 7
AND       P00008	// S_PS_8 Proximity sensor No. 8
AND NOT   P00009	// S_PS_9 Proximity sensor No. 9
MOV       10 D00063	// 중간_빈공간_XGPM Middle empty space XGPM
MLOAD
AND       P00001	// S_PS_1 Proximity sensor No. 1
AND       P00002	// S_PS_2 Proximity sensor No. 2
AND       P00003	// S_PS_3 Proximity sensor No. 3
AND       P00004	// S_PS_4 Proximity sensor No. 4
AND       P00005	// S_PS_5 Proximity sensor No. 5
AND       P00006	// S_PS_6 Proximity sensor No. 6
AND       P00007	// S_PS_7 Proximity sensor No. 7
AND NOT   P00008	// S_PS_8 Proximity sensor No. 8
AND       P00009	// S_PS_9 Proximity sensor No. 9
MOV       9 D00063	// 중간_빈공간_XGPM Middle empty space XGPM
MLOAD
AND       P00001	// S_PS_1 Proximity sensor No. 1
AND       P00002	// S_PS_2 Proximity sensor No. 2
AND       P00003	// S_PS_3 Proximity sensor No. 3
AND       P00004	// S_PS_4 Proximity sensor No. 4
AND       P00005	// S_PS_5 Proximity sensor No. 5
AND       P00006	// S_PS_6 Proximity sensor No. 6
AND NOT   P00007	// S_PS_7 Proximity sensor No. 7
AND       P00008	// S_PS_8 Proximity sensor No. 8
AND       P00009	// S_PS_9 Proximity sensor No. 9
MOV       8 D00063	// 중간_빈공간_XGPM Middle empty space XGPM
MLOAD
AND       P00001	// S_PS_1 Proximity sensor No. 1
AND       P00002	// S_PS_2 Proximity sensor No. 2
AND       P00003	// S_PS_3 Proximity sensor No. 3
AND       P00004	// S_PS_4 Proximity sensor No. 4
AND       P00005	// S_PS_5 Proximity sensor No. 5
AND NOT   P00006	// S_PS_6 Proximity sensor No. 6
AND       P00007	// S_PS_7 Proximity sensor No. 7
AND       P00008	// S_PS_8 Proximity sensor No. 8
AND       P00009	// S_PS_9 Proximity sensor No. 9
MOV       7 D00063	// 중간_빈공간_XGPM Middle empty space XGPM
MLOAD
AND       P00001	// S_PS_1 Proximity sensor No. 1
AND       P00002	// S_PS_2 Proximity sensor No. 2
AND       P00003	// S_PS_3 Proximity sensor No. 3
AND       P00004	// S_PS_4 Proximity sensor No. 4
AND NOT   P00005	// S_PS_5 Proximity sensor No. 5
AND       P00006	// S_PS_6 Proximity sensor No. 6
AND       P00007	// S_PS_7 Proximity sensor No. 7
AND       P00008	// S_PS_8 Proximity sensor No. 8
AND       P00009	// S_PS_9 Proximity sensor No. 9
MOV       6 D00063	// 중간_빈공간_XGPM Middle empty space XGPM
MLOAD
AND       P00001	// S_PS_1 Proximity sensor No. 1
AND       P00002	// S_PS_2 Proximity sensor No. 2
AND       P00003	// S_PS_3 Proximity sensor No. 3
AND NOT   P00004	// S_PS_4 Proximity sensor No. 4
AND       P00005	// S_PS_5 Proximity sensor No. 5
AND       P00006	// S_PS_6 Proximity sensor No. 6
AND       P00007	// S_PS_7 Proximity sensor No. 7
AND       P00008	// S_PS_8 Proximity sensor No. 8
AND       P00009	// S_PS_9 Proximity sensor No. 9
MOV       5 D00063	// 중간_빈공간_XGPM Middle empty space XGPM
MLOAD
AND       P00001	// S_PS_1 Proximity sensor No. 1
AND       P00002	// S_PS_2 Proximity sensor No. 2
AND NOT   P00003	// S_PS_3 Proximity sensor No. 3
AND       P00004	// S_PS_4 Proximity sensor No. 4
AND       P00005	// S_PS_5 Proximity sensor No. 5
AND       P00006	// S_PS_6 Proximity sensor No. 6
AND       P00007	// S_PS_7 Proximity sensor No. 7
AND       P00008	// S_PS_8 Proximity sensor No. 8
AND       P00009	// S_PS_9 Proximity sensor No. 9
MOV       4 D00063	// 중간_빈공간_XGPM Middle empty space XGPM
MLOAD
AND       P00001	// S_PS_1 Proximity sensor No. 1
AND NOT   P00002	// S_PS_2 Proximity sensor No. 2
AND       P00003	// S_PS_3 Proximity sensor No. 3
AND       P00004	// S_PS_4 Proximity sensor No. 4
AND       P00005	// S_PS_5 Proximity sensor No. 5
AND       P00006	// S_PS_6 Proximity sensor No. 6
AND       P00007	// S_PS_7 Proximity sensor No. 7
AND       P00008	// S_PS_8 Proximity sensor No. 8
AND       P00009	// S_PS_9 Proximity sensor No. 9
MOV       3 D00063	// 중간_빈공간_XGPM Middle empty space XGPM
MPOP
AND NOT   P00001	// S_PS_1 Proximity sensor No. 1
AND       P00002	// S_PS_2 Proximity sensor No. 2
AND       P00003	// S_PS_3 Proximity sensor No. 3
AND       P00004	// S_PS_4 Proximity sensor No. 4
AND       P00005	// S_PS_5 Proximity sensor No. 5
AND       P00006	// S_PS_6 Proximity sensor No. 6
AND       P00007	// S_PS_7 Proximity sensor No. 7
AND       P00008	// S_PS_8 Proximity sensor No. 8
AND       P00009	// S_PS_9 Proximity sensor No. 9
MOV       2 D00063	// 중간_빈공간_XGPM Middle empty space XGPM

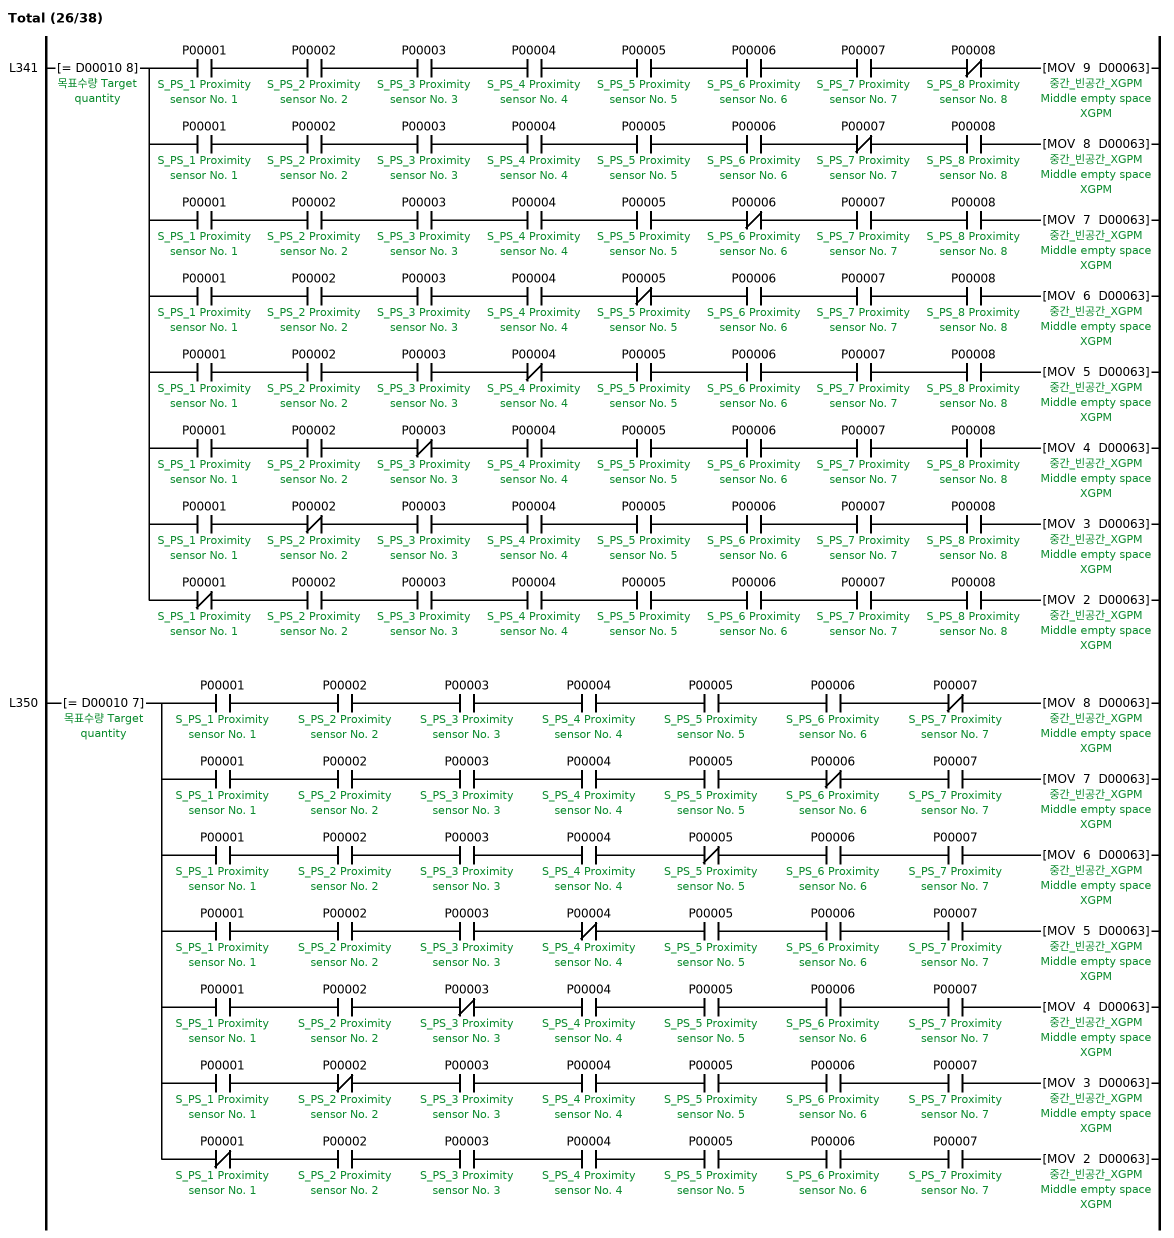
; L341
LOAD=     D00010 8	// 목표수량 Target quantity
MPUSH
AND       P00001	// S_PS_1 Proximity sensor No. 1
AND       P00002	// S_PS_2 Proximity sensor No. 2
AND       P00003	// S_PS_3 Proximity sensor No. 3
AND       P00004	// S_PS_4 Proximity sensor No. 4
AND       P00005	// S_PS_5 Proximity sensor No. 5
AND       P00006	// S_PS_6 Proximity sensor No. 6
AND       P00007	// S_PS_7 Proximity sensor No. 7
AND NOT   P00008	// S_PS_8 Proximity sensor No. 8
MOV       9 D00063	// 중간_빈공간_XGPM Middle empty space XGPM
MLOAD
AND       P00001	// S_PS_1 Proximity sensor No. 1
AND       P00002	// S_PS_2 Proximity sensor No. 2
AND       P00003	// S_PS_3 Proximity sensor No. 3
AND       P00004	// S_PS_4 Proximity sensor No. 4
AND       P00005	// S_PS_5 Proximity sensor No. 5
AND       P00006	// S_PS_6 Proximity sensor No. 6
AND NOT   P00007	// S_PS_7 Proximity sensor No. 7
AND       P00008	// S_PS_8 Proximity sensor No. 8
MOV       8 D00063	// 중간_빈공간_XGPM Middle empty space XGPM
MLOAD
AND       P00001	// S_PS_1 Proximity sensor No. 1
AND       P00002	// S_PS_2 Proximity sensor No. 2
AND       P00003	// S_PS_3 Proximity sensor No. 3
AND       P00004	// S_PS_4 Proximity sensor No. 4
AND       P00005	// S_PS_5 Proximity sensor No. 5
AND NOT   P00006	// S_PS_6 Proximity sensor No. 6
AND       P00007	// S_PS_7 Proximity sensor No. 7
AND       P00008	// S_PS_8 Proximity sensor No. 8
MOV       7 D00063	// 중간_빈공간_XGPM Middle empty space XGPM
MLOAD
AND       P00001	// S_PS_1 Proximity sensor No. 1
AND       P00002	// S_PS_2 Proximity sensor No. 2
AND       P00003	// S_PS_3 Proximity sensor No. 3
AND       P00004	// S_PS_4 Proximity sensor No. 4
AND NOT   P00005	// S_PS_5 Proximity sensor No. 5
AND       P00006	// S_PS_6 Proximity sensor No. 6
AND       P00007	// S_PS_7 Proximity sensor No. 7
AND       P00008	// S_PS_8 Proximity sensor No. 8
MOV       6 D00063	// 중간_빈공간_XGPM Middle empty space XGPM
MLOAD
AND       P00001	// S_PS_1 Proximity sensor No. 1
AND       P00002	// S_PS_2 Proximity sensor No. 2
AND       P00003	// S_PS_3 Proximity sensor No. 3
AND NOT   P00004	// S_PS_4 Proximity sensor No. 4
AND       P00005	// S_PS_5 Proximity sensor No. 5
AND       P00006	// S_PS_6 Proximity sensor No. 6
AND       P00007	// S_PS_7 Proximity sensor No. 7
AND       P00008	// S_PS_8 Proximity sensor No. 8
MOV       5 D00063	// 중간_빈공간_XGPM Middle empty space XGPM
MLOAD
AND       P00001	// S_PS_1 Proximity sensor No. 1
AND       P00002	// S_PS_2 Proximity sensor No. 2
AND NOT   P00003	// S_PS_3 Proximity sensor No. 3
AND       P00004	// S_PS_4 Proximity sensor No. 4
AND       P00005	// S_PS_5 Proximity sensor No. 5
AND       P00006	// S_PS_6 Proximity sensor No. 6
AND       P00007	// S_PS_7 Proximity sensor No. 7
AND       P00008	// S_PS_8 Proximity sensor No. 8
MOV       4 D00063	// 중간_빈공간_XGPM Middle empty space XGPM
MLOAD
AND       P00001	// S_PS_1 Proximity sensor No. 1
AND NOT   P00002	// S_PS_2 Proximity sensor No. 2
AND       P00003	// S_PS_3 Proximity sensor No. 3
AND       P00004	// S_PS_4 Proximity sensor No. 4
AND       P00005	// S_PS_5 Proximity sensor No. 5
AND       P00006	// S_PS_6 Proximity sensor No. 6
AND       P00007	// S_PS_7 Proximity sensor No. 7
AND       P00008	// S_PS_8 Proximity sensor No. 8
MOV       3 D00063	// 중간_빈공간_XGPM Middle empty space XGPM
MPOP
AND NOT   P00001	// S_PS_1 Proximity sensor No. 1
AND       P00002	// S_PS_2 Proximity sensor No. 2
AND       P00003	// S_PS_3 Proximity sensor No. 3
AND       P00004	// S_PS_4 Proximity sensor No. 4
AND       P00005	// S_PS_5 Proximity sensor No. 5
AND       P00006	// S_PS_6 Proximity sensor No. 6
AND       P00007	// S_PS_7 Proximity sensor No. 7
AND       P00008	// S_PS_8 Proximity sensor No. 8
MOV       2 D00063	// 중간_빈공간_XGPM Middle empty space XGPM
; L350
LOAD=     D00010 7	// 목표수량 Target quantity
MPUSH
AND       P00001	// S_PS_1 Proximity sensor No. 1
AND       P00002	// S_PS_2 Proximity sensor No. 2
AND       P00003	// S_PS_3 Proximity sensor No. 3
AND       P00004	// S_PS_4 Proximity sensor No. 4
AND       P00005	// S_PS_5 Proximity sensor No. 5
AND       P00006	// S_PS_6 Proximity sensor No. 6
AND NOT   P00007	// S_PS_7 Proximity sensor No. 7
MOV       8 D00063	// 중간_빈공간_XGPM Middle empty space XGPM
MLOAD
AND       P00001	// S_PS_1 Proximity sensor No. 1
AND       P00002	// S_PS_2 Proximity sensor No. 2
AND       P00003	// S_PS_3 Proximity sensor No. 3
AND       P00004	// S_PS_4 Proximity sensor No. 4
AND       P00005	// S_PS_5 Proximity sensor No. 5
AND NOT   P00006	// S_PS_6 Proximity sensor No. 6
AND       P00007	// S_PS_7 Proximity sensor No. 7
MOV       7 D00063	// 중간_빈공간_XGPM Middle empty space XGPM
MLOAD
AND       P00001	// S_PS_1 Proximity sensor No. 1
AND       P00002	// S_PS_2 Proximity sensor No. 2
AND       P00003	// S_PS_3 Proximity sensor No. 3
AND       P00004	// S_PS_4 Proximity sensor No. 4
AND NOT   P00005	// S_PS_5 Proximity sensor No. 5
AND       P00006	// S_PS_6 Proximity sensor No. 6
AND       P00007	// S_PS_7 Proximity sensor No. 7
MOV       6 D00063	// 중간_빈공간_XGPM Middle empty space XGPM
MLOAD
AND       P00001	// S_PS_1 Proximity sensor No. 1
AND       P00002	// S_PS_2 Proximity sensor No. 2
AND       P00003	// S_PS_3 Proximity sensor No. 3
AND NOT   P00004	// S_PS_4 Proximity sensor No. 4
AND       P00005	// S_PS_5 Proximity sensor No. 5
AND       P00006	// S_PS_6 Proximity sensor No. 6
AND       P00007	// S_PS_7 Proximity sensor No. 7
MOV       5 D00063	// 중간_빈공간_XGPM Middle empty space XGPM
MLOAD
AND       P00001	// S_PS_1 Proximity sensor No. 1
AND       P00002	// S_PS_2 Proximity sensor No. 2
AND NOT   P00003	// S_PS_3 Proximity sensor No. 3
AND       P00004	// S_PS_4 Proximity sensor No. 4
AND       P00005	// S_PS_5 Proximity sensor No. 5
AND       P00006	// S_PS_6 Proximity sensor No. 6
AND       P00007	// S_PS_7 Proximity sensor No. 7
MOV       4 D00063	// 중간_빈공간_XGPM Middle empty space XGPM
MLOAD
AND       P00001	// S_PS_1 Proximity sensor No. 1
AND NOT   P00002	// S_PS_2 Proximity sensor No. 2
AND       P00003	// S_PS_3 Proximity sensor No. 3
AND       P00004	// S_PS_4 Proximity sensor No. 4
AND       P00005	// S_PS_5 Proximity sensor No. 5
AND       P00006	// S_PS_6 Proximity sensor No. 6
AND       P00007	// S_PS_7 Proximity sensor No. 7
MOV       3 D00063	// 중간_빈공간_XGPM Middle empty space XGPM
MPOP
AND NOT   P00001	// S_PS_1 Proximity sensor No. 1
AND       P00002	// S_PS_2 Proximity sensor No. 2
AND       P00003	// S_PS_3 Proximity sensor No. 3
AND       P00004	// S_PS_4 Proximity sensor No. 4
AND       P00005	// S_PS_5 Proximity sensor No. 5
AND       P00006	// S_PS_6 Proximity sensor No. 6
AND       P00007	// S_PS_7 Proximity sensor No. 7
MOV       2 D00063	// 중간_빈공간_XGPM Middle empty space XGPM

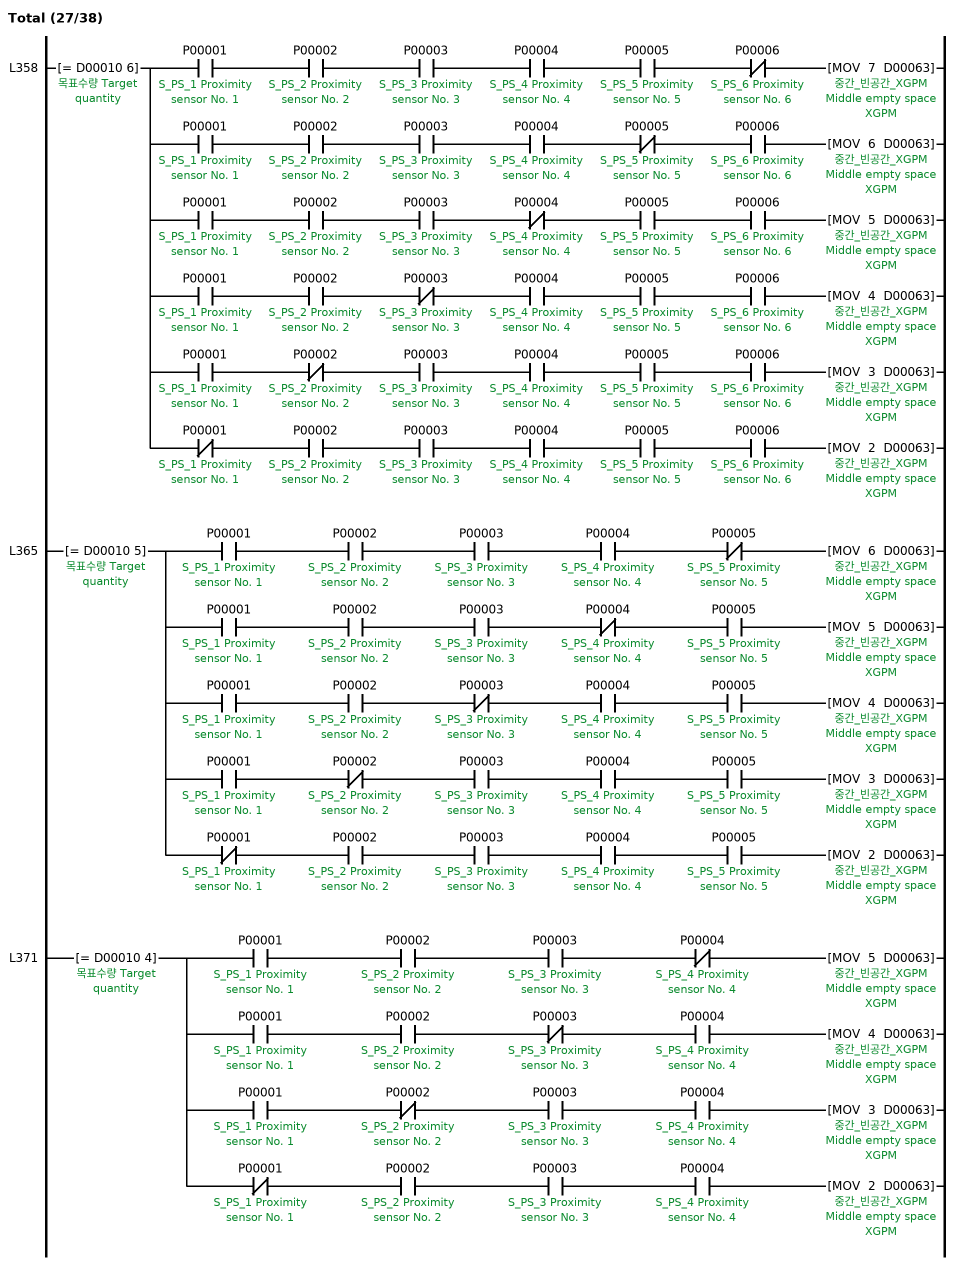
; L358
LOAD=     D00010 6	// 목표수량 Target quantity
MPUSH
AND       P00001	// S_PS_1 Proximity sensor No. 1
AND       P00002	// S_PS_2 Proximity sensor No. 2
AND       P00003	// S_PS_3 Proximity sensor No. 3
AND       P00004	// S_PS_4 Proximity sensor No. 4
AND       P00005	// S_PS_5 Proximity sensor No. 5
AND NOT   P00006	// S_PS_6 Proximity sensor No. 6
MOV       7 D00063	// 중간_빈공간_XGPM Middle empty space XGPM
MLOAD
AND       P00001	// S_PS_1 Proximity sensor No. 1
AND       P00002	// S_PS_2 Proximity sensor No. 2
AND       P00003	// S_PS_3 Proximity sensor No. 3
AND       P00004	// S_PS_4 Proximity sensor No. 4
AND NOT   P00005	// S_PS_5 Proximity sensor No. 5
AND       P00006	// S_PS_6 Proximity sensor No. 6
MOV       6 D00063	// 중간_빈공간_XGPM Middle empty space XGPM
MLOAD
AND       P00001	// S_PS_1 Proximity sensor No. 1
AND       P00002	// S_PS_2 Proximity sensor No. 2
AND       P00003	// S_PS_3 Proximity sensor No. 3
AND NOT   P00004	// S_PS_4 Proximity sensor No. 4
AND       P00005	// S_PS_5 Proximity sensor No. 5
AND       P00006	// S_PS_6 Proximity sensor No. 6
MOV       5 D00063	// 중간_빈공간_XGPM Middle empty space XGPM
MLOAD
AND       P00001	// S_PS_1 Proximity sensor No. 1
AND       P00002	// S_PS_2 Proximity sensor No. 2
AND NOT   P00003	// S_PS_3 Proximity sensor No. 3
AND       P00004	// S_PS_4 Proximity sensor No. 4
AND       P00005	// S_PS_5 Proximity sensor No. 5
AND       P00006	// S_PS_6 Proximity sensor No. 6
MOV       4 D00063	// 중간_빈공간_XGPM Middle empty space XGPM
MLOAD
AND       P00001	// S_PS_1 Proximity sensor No. 1
AND NOT   P00002	// S_PS_2 Proximity sensor No. 2
AND       P00003	// S_PS_3 Proximity sensor No. 3
AND       P00004	// S_PS_4 Proximity sensor No. 4
AND       P00005	// S_PS_5 Proximity sensor No. 5
AND       P00006	// S_PS_6 Proximity sensor No. 6
MOV       3 D00063	// 중간_빈공간_XGPM Middle empty space XGPM
MPOP
AND NOT   P00001	// S_PS_1 Proximity sensor No. 1
AND       P00002	// S_PS_2 Proximity sensor No. 2
AND       P00003	// S_PS_3 Proximity sensor No. 3
AND       P00004	// S_PS_4 Proximity sensor No. 4
AND       P00005	// S_PS_5 Proximity sensor No. 5
AND       P00006	// S_PS_6 Proximity sensor No. 6
MOV       2 D00063	// 중간_빈공간_XGPM Middle empty space XGPM
; L365
LOAD=     D00010 5	// 목표수량 Target quantity
MPUSH
AND       P00001	// S_PS_1 Proximity sensor No. 1
AND       P00002	// S_PS_2 Proximity sensor No. 2
AND       P00003	// S_PS_3 Proximity sensor No. 3
AND       P00004	// S_PS_4 Proximity sensor No. 4
AND NOT   P00005	// S_PS_5 Proximity sensor No. 5
MOV       6 D00063	// 중간_빈공간_XGPM Middle empty space XGPM
MLOAD
AND       P00001	// S_PS_1 Proximity sensor No. 1
AND       P00002	// S_PS_2 Proximity sensor No. 2
AND       P00003	// S_PS_3 Proximity sensor No. 3
AND NOT   P00004	// S_PS_4 Proximity sensor No. 4
AND       P00005	// S_PS_5 Proximity sensor No. 5
MOV       5 D00063	// 중간_빈공간_XGPM Middle empty space XGPM
MLOAD
AND       P00001	// S_PS_1 Proximity sensor No. 1
AND       P00002	// S_PS_2 Proximity sensor No. 2
AND NOT   P00003	// S_PS_3 Proximity sensor No. 3
AND       P00004	// S_PS_4 Proximity sensor No. 4
AND       P00005	// S_PS_5 Proximity sensor No. 5
MOV       4 D00063	// 중간_빈공간_XGPM Middle empty space XGPM
MLOAD
AND       P00001	// S_PS_1 Proximity sensor No. 1
AND NOT   P00002	// S_PS_2 Proximity sensor No. 2
AND       P00003	// S_PS_3 Proximity sensor No. 3
AND       P00004	// S_PS_4 Proximity sensor No. 4
AND       P00005	// S_PS_5 Proximity sensor No. 5
MOV       3 D00063	// 중간_빈공간_XGPM Middle empty space XGPM
MPOP
AND NOT   P00001	// S_PS_1 Proximity sensor No. 1
AND       P00002	// S_PS_2 Proximity sensor No. 2
AND       P00003	// S_PS_3 Proximity sensor No. 3
AND       P00004	// S_PS_4 Proximity sensor No. 4
AND       P00005	// S_PS_5 Proximity sensor No. 5
MOV       2 D00063	// 중간_빈공간_XGPM Middle empty space XGPM
; L371
LOAD=     D00010 4	// 목표수량 Target quantity
MPUSH
AND       P00001	// S_PS_1 Proximity sensor No. 1
AND       P00002	// S_PS_2 Proximity sensor No. 2
AND       P00003	// S_PS_3 Proximity sensor No. 3
AND NOT   P00004	// S_PS_4 Proximity sensor No. 4
MOV       5 D00063	// 중간_빈공간_XGPM Middle empty space XGPM
MLOAD
AND       P00001	// S_PS_1 Proximity sensor No. 1
AND       P00002	// S_PS_2 Proximity sensor No. 2
AND NOT   P00003	// S_PS_3 Proximity sensor No. 3
AND       P00004	// S_PS_4 Proximity sensor No. 4
MOV       4 D00063	// 중간_빈공간_XGPM Middle empty space XGPM
MLOAD
AND       P00001	// S_PS_1 Proximity sensor No. 1
AND NOT   P00002	// S_PS_2 Proximity sensor No. 2
AND       P00003	// S_PS_3 Proximity sensor No. 3
AND       P00004	// S_PS_4 Proximity sensor No. 4
MOV       3 D00063	// 중간_빈공간_XGPM Middle empty space XGPM
MPOP
AND NOT   P00001	// S_PS_1 Proximity sensor No. 1
AND       P00002	// S_PS_2 Proximity sensor No. 2
AND       P00003	// S_PS_3 Proximity sensor No. 3
AND       P00004	// S_PS_4 Proximity sensor No. 4
MOV       2 D00063	// 중간_빈공간_XGPM Middle empty space XGPM

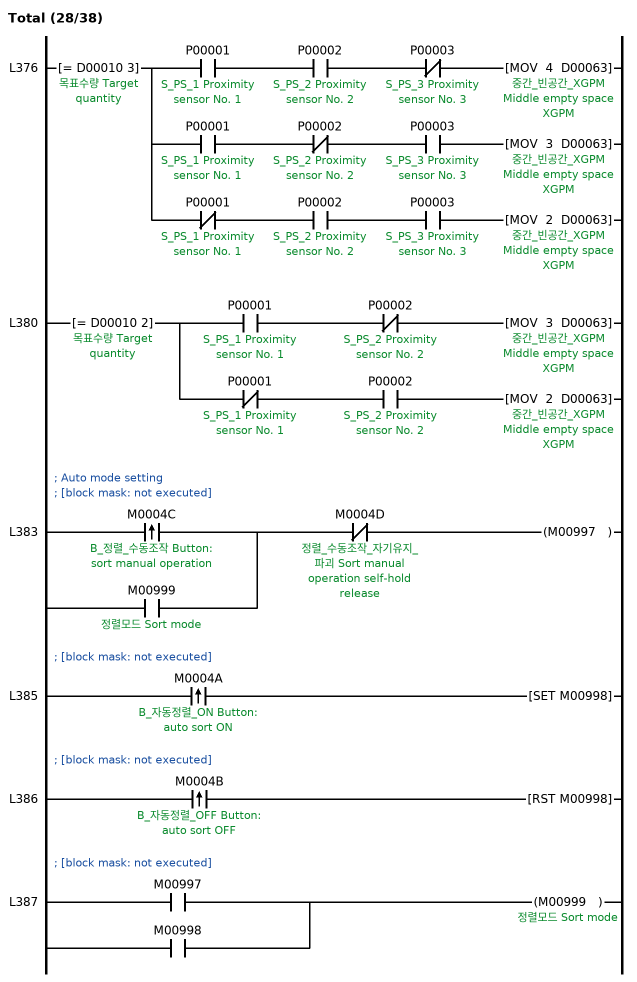
; L376
LOAD=     D00010 3	// 목표수량 Target quantity
MPUSH
AND       P00001	// S_PS_1 Proximity sensor No. 1
AND       P00002	// S_PS_2 Proximity sensor No. 2
AND NOT   P00003	// S_PS_3 Proximity sensor No. 3
MOV       4 D00063	// 중간_빈공간_XGPM Middle empty space XGPM
MLOAD
AND       P00001	// S_PS_1 Proximity sensor No. 1
AND NOT   P00002	// S_PS_2 Proximity sensor No. 2
AND       P00003	// S_PS_3 Proximity sensor No. 3
MOV       3 D00063	// 중간_빈공간_XGPM Middle empty space XGPM
MPOP
AND NOT   P00001	// S_PS_1 Proximity sensor No. 1
AND       P00002	// S_PS_2 Proximity sensor No. 2
AND       P00003	// S_PS_3 Proximity sensor No. 3
MOV       2 D00063	// 중간_빈공간_XGPM Middle empty space XGPM
; L380
LOAD=     D00010 2	// 목표수량 Target quantity
MPUSH
AND       P00001	// S_PS_1 Proximity sensor No. 1
AND NOT   P00002	// S_PS_2 Proximity sensor No. 2
MOV       3 D00063	// 중간_빈공간_XGPM Middle empty space XGPM
MPOP
AND NOT   P00001	// S_PS_1 Proximity sensor No. 1
AND       P00002	// S_PS_2 Proximity sensor No. 2
MOV       2 D00063	// 중간_빈공간_XGPM Middle empty space XGPM
// Auto mode setting
; L383 (block mask: not executed)
LOADP     M0004C	// B_정렬_수동조작 Button: sort manual operation
OR        M00999	// 정렬모드 Sort mode
AND NOT   M0004D	// 정렬_수동조작_자기유지_파괴 Sort manual operation self-hold release
OUT       M00997
; L385 (block mask: not executed)
LOADP     M0004A	// B_자동정렬_ON Button: auto sort ON
SET       M00998
; L386 (block mask: not executed)
LOADP     M0004B	// B_자동정렬_OFF Button: auto sort OFF
RST       M00998
; L387 (block mask: not executed)
LOAD      M00997
OR        M00998
OUT       M00999	// 정렬모드 Sort mode

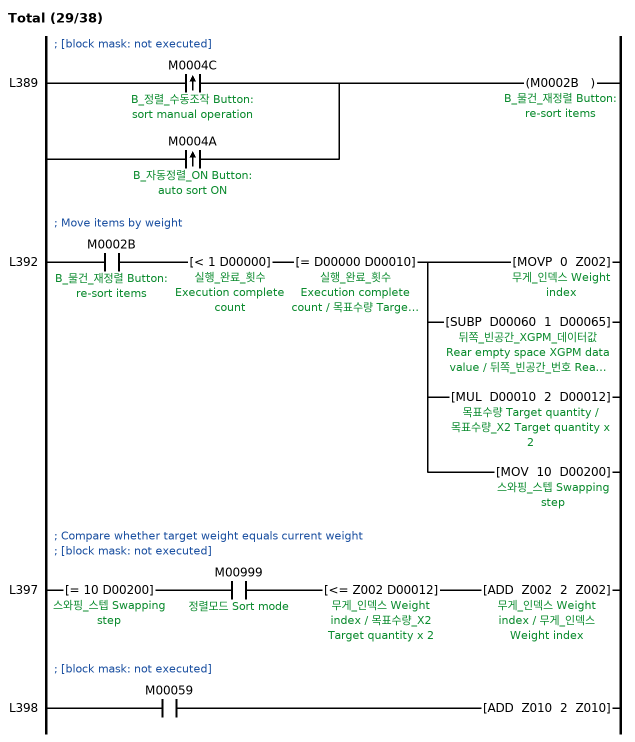
; L389 (block mask: not executed)
LOADP     M0004C	// B_정렬_수동조작 Button: sort manual operation
ORP       M0004A	// B_자동정렬_ON Button: auto sort ON
OUT       M0002B	// B_물건_재정렬 Button: re-sort items
// Move items by weight
; L392
LOAD      M0002B	// B_물건_재정렬 Button: re-sort items
AND<      1 D00000	// 실행_완료_횟수 Execution complete count
AND=      D00000 D00010	// 실행_완료_횟수 Execution complete count / 목표수량 Target quantity
MOVP      0 Z002	// 무게_인덱스 Weight index
SUBP      D00060 1 D00065	// 뒤쪽_빈공간_XGPM_데이터값 Rear empty space XGPM data value / 뒤쪽_빈공간_번호 Rear empty space number
MUL       D00010 2 D00012	// 목표수량 Target quantity / 목표수량_X2 Target quantity x 2
MOV       10 D00200	// 스와핑_스텝 Swapping step
// Compare whether target weight equals current weight
; L397 (block mask: not executed)
LOAD=     10 D00200	// 스와핑_스텝 Swapping step
AND       M00999	// 정렬모드 Sort mode
AND<=     Z002 D00012	// 무게_인덱스 Weight index / 목표수량_X2 Target quantity x 2
ADD       Z002 2 Z002	// 무게_인덱스 Weight index / 무게_인덱스 Weight index
; L398 (block mask: not executed)
LOAD      M00059
ADD       Z010 2 Z010

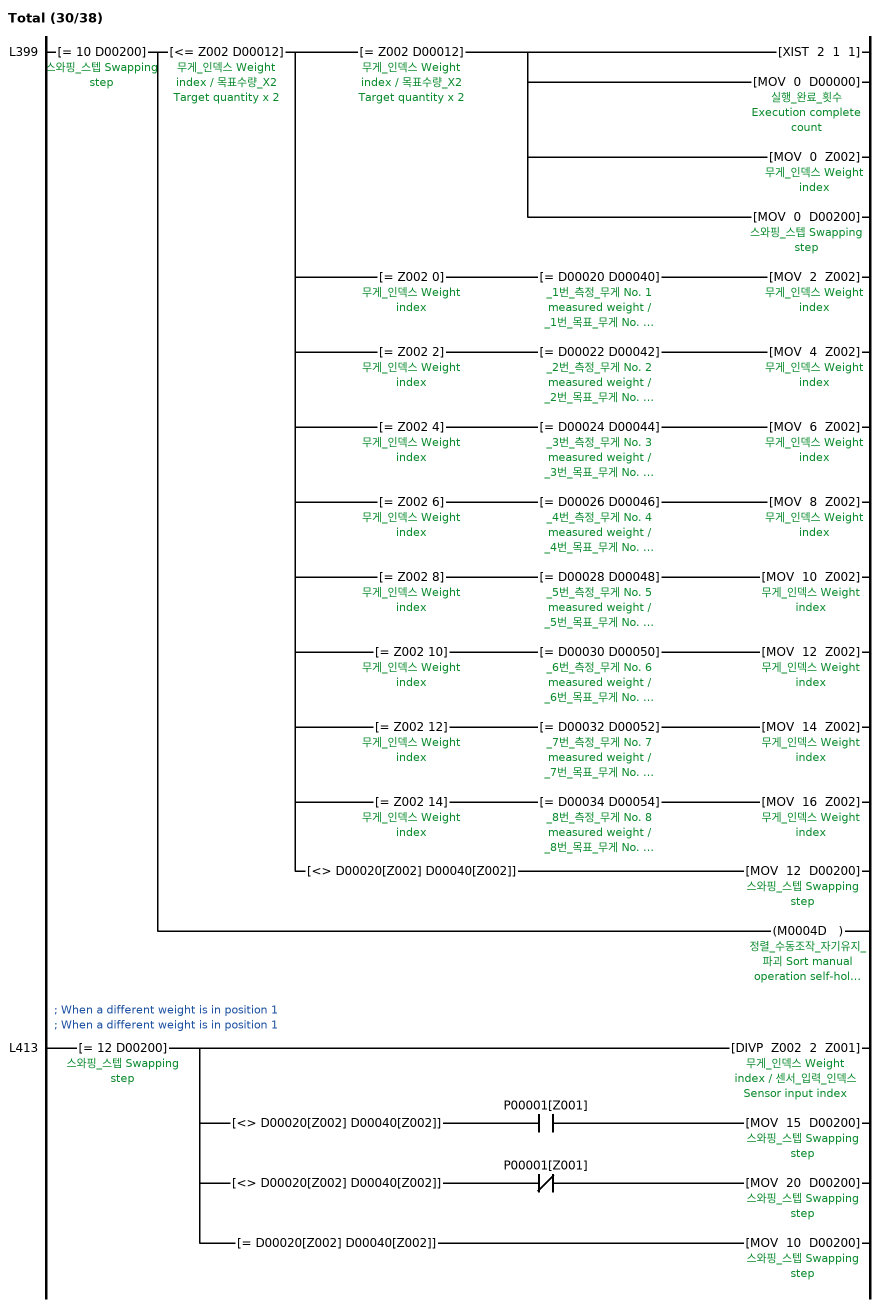
; L399
LOAD=     10 D00200	// 스와핑_스텝 Swapping step
MPUSH
AND<=     Z002 D00012	// 무게_인덱스 Weight index / 목표수량_X2 Target quantity x 2
MPUSH
AND=      Z002 D00012	// 무게_인덱스 Weight index / 목표수량_X2 Target quantity x 2
XIST      2 1 1
MOV       0 D00000	// 실행_완료_횟수 Execution complete count
MOV       0 Z002	// 무게_인덱스 Weight index
MOV       0 D00200	// 스와핑_스텝 Swapping step
MLOAD
AND=      Z002 0	// 무게_인덱스 Weight index
AND=      D00020 D00040	// _1번_측정_무게 No. 1 measured weight / _1번_목표_무게 No. 1 target weight
MOV       2 Z002	// 무게_인덱스 Weight index
MLOAD
AND=      Z002 2	// 무게_인덱스 Weight index
AND=      D00022 D00042	// _2번_측정_무게 No. 2 measured weight / _2번_목표_무게 No. 2 target weight
MOV       4 Z002	// 무게_인덱스 Weight index
MLOAD
AND=      Z002 4	// 무게_인덱스 Weight index
AND=      D00024 D00044	// _3번_측정_무게 No. 3 measured weight / _3번_목표_무게 No. 3 target weight
MOV       6 Z002	// 무게_인덱스 Weight index
MLOAD
AND=      Z002 6	// 무게_인덱스 Weight index
AND=      D00026 D00046	// _4번_측정_무게 No. 4 measured weight / _4번_목표_무게 No. 4 target weight
MOV       8 Z002	// 무게_인덱스 Weight index
MLOAD
AND=      Z002 8	// 무게_인덱스 Weight index
AND=      D00028 D00048	// _5번_측정_무게 No. 5 measured weight / _5번_목표_무게 No. 5 target weight
MOV       10 Z002	// 무게_인덱스 Weight index
MLOAD
AND=      Z002 10	// 무게_인덱스 Weight index
AND=      D00030 D00050	// _6번_측정_무게 No. 6 measured weight / _6번_목표_무게 No. 6 target weight
MOV       12 Z002	// 무게_인덱스 Weight index
MLOAD
AND=      Z002 12	// 무게_인덱스 Weight index
AND=      D00032 D00052	// _7번_측정_무게 No. 7 measured weight / _7번_목표_무게 No. 7 target weight
MOV       14 Z002	// 무게_인덱스 Weight index
MLOAD
AND=      Z002 14	// 무게_인덱스 Weight index
AND=      D00034 D00054	// _8번_측정_무게 No. 8 measured weight / _8번_목표_무게 No. 8 target weight
MOV       16 Z002	// 무게_인덱스 Weight index
MPOP
AND<>     D00020[Z002] D00040[Z002]
MOV       12 D00200	// 스와핑_스텝 Swapping step
MPOP
OUT       M0004D	// 정렬_수동조작_자기유지_파괴 Sort manual operation self-hold release
; L413
LOAD=     12 D00200	// 스와핑_스텝 Swapping step
DIVP      Z002 2 Z001	// 무게_인덱스 Weight index / 센서_입력_인덱스 Sensor input index
MPUSH
AND<>     D00020[Z002] D00040[Z002]
AND       P00001[Z001]
MOV       15 D00200	// 스와핑_스텝 Swapping step
MLOAD
AND<>     D00020[Z002] D00040[Z002]
AND NOT   P00001[Z001]
MOV       20 D00200	// 스와핑_스텝 Swapping step
MPOP
AND=      D00020[Z002] D00040[Z002]
MOV       10 D00200	// 스와핑_스텝 Swapping step
// output comment: When a different weight is in position 1
// output comment: When a different weight is in position 1

